--- program cerlaizgr (robot Fanuc LR Mate 200iD/7L) ---
  Suave(1)
  Establecer velocidad (1000.0 mm/s)
  Est. Ref.: bote cera
  Est. herr: Tool 1
  Mostrar Tool 1
  MoveJ 1 to (318.69, -45.69, 237.74) mm, rotated rx 168.3 ry -14.7 rz -86.98 deg; joints [83.928, 45.745, -7.693, -16.831, -73.362, 101.148]
  MoveL 2 to (318.69, -45.69, 237.74) mm, rotated rx 168.3 ry -14.7 rz -86.98 deg; joints [83.928, 45.745, -7.693, -16.831, -73.362, 101.148]
  MoveL 3 to (299.08, -45.69, 139.68) mm, rotated rx 168.3 ry -14.7 rz -86.98 deg; joints [84.076, 51.288, -16.777, -17.851, -64.646, 103.898]
  MoveL 4 to (299.08, -45.69, 139.68) mm, rotated rx 168.3 ry -14.7 rz -86.98 deg; joints [84.076, 51.288, -16.777, -17.851, -64.646, 103.898]
  Establecer velocidad (50.0 mm/s)
  MoveL 5 to (313.16, -44.5, 139.68) mm, rotated rx 168.3 ry -14.7 rz -86.98 deg; joints [83.886, 49.076, -18.597, -18.155, -62.971, 104.717]
  MoveL 6 to (327.32, -44.52, 139.68) mm, rotated rx 168.3 ry -14.7 rz -86.98 deg; joints [83.776, 46.952, -20.301, -18.453, -61.386, 105.433]
  MoveL 7 to (341.43, -45.73, 139.68) mm, rotated rx 168.3 ry -14.7 rz -86.98 deg; joints [83.752, 44.917, -21.892, -18.741, -59.886, 106.039]
  MoveL 8 to (355.34, -48.13, 139.68) mm, rotated rx 168.3 ry -14.7 rz -86.98 deg; joints [83.819, 42.973, -23.371, -19.018, -58.466, 106.529]
  MoveL 9 to (368.95, -51.69, 140.34) mm, rotated rx 168.3 ry -14.7 rz -86.98 deg; joints [83.98, 41.087, -24.673, -19.265, -57.187, 106.869]
  MoveL 10 to (383, -56.41, 142.33) mm, rotated rx 168.3 ry -14.7 rz -86.98 deg; joints [84.236, 39.118, -25.797, -19.475, -56.051, 107.053]
  MoveL 11 to (396.92, -60.57, 145.69) mm, rotated rx 168.3 ry -14.7 rz -86.98 deg; joints [84.459, 37.148, -26.671, -19.645, -55.16, 107.18]
  MoveL 12 to (410.7, -63.96, 150.39) mm, rotated rx 168.3 ry -14.7 rz -86.98 deg; joints [84.628, 35.164, -27.3, -19.771, -54.517, 107.266]
  MoveL 13 to (424.7, -66.68, 154.58) mm, rotated rx 168.3 ry -14.7 rz -86.98 deg; joints [84.746, 33.212, -27.925, -19.908, -53.893, 107.406]
  MoveL 14 to (439.04, -68.74, 157.38) mm, rotated rx 168.3 ry -14.7 rz -86.98 deg; joints [84.81, 31.317, -28.662, -20.086, -53.182, 107.653]
  MoveL 15 to (453.73, -70.09, 158.77) mm, rotated rx 168.3 ry -14.7 rz -86.98 deg; joints [84.812, 29.481, -29.518, -20.31, -52.377, 108.022]
  MoveL 16 to (469.71, -70.72, 158.92) mm, rotated rx 168.3 ry -14.7 rz -86.98 deg; joints [84.738, 27.589, -30.539, -20.6, -51.443, 108.552]
  MoveL 17 to (485.71, -70.47, 158.92) mm, rotated rx 168.3 ry -14.7 rz -86.98 deg; joints [84.58, 25.732, -31.509, -20.899, -50.584, 109.158]
  MoveL 18 to (501.7, -70.47, 158.92) mm, rotated rx 168.3 ry -14.7 rz -86.98 deg; joints [84.436, 23.886, -32.418, -21.19, -49.78, 109.731]
  MoveL 19 to (517.7, -70.47, 158.92) mm, rotated rx 168.3 ry -14.7 rz -86.98 deg; joints [84.284, 22.05, -33.266, -21.473, -49.036, 110.293]
  MoveL 20 to (533.69, -70.47, 158.92) mm, rotated rx 168.3 ry -14.7 rz -86.98 deg; joints [84.125, 20.219, -34.053, -21.748, -48.354, 110.844]
  MoveL 21 to (543.69, -70.47, 158.92) mm, rotated rx 168.3 ry -14.7 rz -86.98 deg; joints [84.02, 19.075, -34.514, -21.915, -47.958, 111.182]
  MoveL 22 to (553.68, -70.47, 158.92) mm, rotated rx 168.3 ry -14.7 rz -86.98 deg; joints [83.912, 17.931, -34.952, -22.077, -47.585, 111.515]
  MoveL 23 to (563.68, -70.47, 158.92) mm, rotated rx 168.3 ry -14.7 rz -86.98 deg; joints [83.799, 16.785, -35.366, -22.234, -47.237, 111.842]
  MoveL 24 to (573.77, -70.76, 158.92) mm, rotated rx 168.3 ry -14.7 rz -86.98 deg; joints [83.713, 15.622, -35.76, -22.383, -46.898, 112.135]
  MoveL 25 to (580.76, -72.49, 158.92) mm, rotated rx 168.3 ry -14.7 rz -86.98 deg; joints [83.817, 14.795, -36.025, -22.466, -46.622, 112.166]
  MoveL 26 to (587.5, -75.89, 158.92) mm, rotated rx 168.3 ry -14.7 rz -86.98 deg; joints [84.112, 13.973, -36.274, -22.521, -46.3, 111.995]
  MoveL 27 to (593.42, -80.86, 158.92) mm, rotated rx 168.3 ry -14.7 rz -86.98 deg; joints [84.6, 13.23, -36.489, -22.541, -45.951, 111.605]
  MoveL 28 to (598, -87.04, 158.92) mm, rotated rx 168.3 ry -14.7 rz -86.98 deg; joints [85.251, 12.632, -36.653, -22.52, -45.6, 111.02]
  MoveL 29 to (600.96, -93.88, 158.92) mm, rotated rx 168.3 ry -14.7 rz -86.98 deg; joints [86.003, 12.225, -36.76, -22.461, -45.269, 110.295]
  MoveL 30 to (602.27, -100.81, 158.92) mm, rotated rx 168.3 ry -14.7 rz -86.98 deg; joints [86.787, 12.02, -36.813, -22.373, -44.981, 109.505]
  MoveL 31 to (602.38, -107.49, 158.92) mm, rotated rx 168.3 ry -14.7 rz -86.98 deg; joints [87.553, 11.969, -36.826, -22.267, -44.736, 108.707]
  MoveL 32 to (602.38, -114.16, 158.92) mm, rotated rx 168.3 ry -14.7 rz -86.98 deg; joints [88.319, 11.941, -36.833, -22.154, -44.498, 107.903]
  MoveL 33 to (601.73, -120.97, 158.92) mm, rotated rx 168.3 ry -14.7 rz -86.98 deg; joints [89.103, 12, -36.818, -22.024, -44.276, 107.063]
  MoveL 34 to (599.51, -127.92, 158.92) mm, rotated rx 168.3 ry -14.7 rz -86.98 deg; joints [89.902, 12.254, -36.753, -21.866, -44.097, 106.177]
  MoveL 35 to (595.62, -134.46, 158.92) mm, rotated rx 168.3 ry -14.7 rz -86.98 deg; joints [90.646, 12.713, -36.63, -21.691, -43.99, 105.315]
  MoveL 36 to (590.24, -140.02, 158.92) mm, rotated rx 168.3 ry -14.7 rz -86.98 deg; joints [91.263, 13.353, -36.453, -21.513, -43.972, 104.557]
  MoveL 37 to (583.78, -144.14, 158.92) mm, rotated rx 168.3 ry -14.7 rz -86.98 deg; joints [91.703, 14.118, -36.231, -21.348, -44.05, 103.965]
  MoveL 38 to (576.83, -146.59, 158.92) mm, rotated rx 168.3 ry -14.7 rz -86.98 deg; joints [91.949, 14.935, -35.98, -21.209, -44.211, 103.569]
  MoveL 39 to (567.71, -147.44, 158.92) mm, rotated rx 168.3 ry -14.7 rz -86.98 deg; joints [92.006, 15.993, -35.636, -21.071, -44.515, 103.329]
  MoveL 40 to (558.83, -147.44, 158.92) mm, rotated rx 168.3 ry -14.7 rz -86.98 deg; joints [91.973, 17.018, -35.283, -20.949, -44.855, 103.185]
  MoveL 41 to (549.94, -147.44, 158.92) mm, rotated rx 168.3 ry -14.7 rz -86.98 deg; joints [91.941, 18.042, -34.91, -20.822, -45.212, 103.031]
  MoveL 42 to (541.06, -147.44, 158.92) mm, rotated rx 168.3 ry -14.7 rz -86.98 deg; joints [91.91, 19.064, -34.518, -20.691, -45.588, 102.87]
  MoveL 43 to (532.17, -147.44, 158.92) mm, rotated rx 168.3 ry -14.7 rz -86.98 deg; joints [91.88, 20.086, -34.107, -20.556, -45.981, 102.7]
  MoveL 44 to (523.28, -147.44, 158.92) mm, rotated rx 168.3 ry -14.7 rz -86.98 deg; joints [91.851, 21.107, -33.678, -20.417, -46.392, 102.523]
  MoveL 45 to (505.69, -147.44, 158.92) mm, rotated rx 168.3 ry -14.7 rz -86.98 deg; joints [91.796, 23.133, -32.772, -20.133, -47.257, 102.152]
  MoveL 46 to (488.1, -147.44, 158.92) mm, rotated rx 168.3 ry -14.7 rz -86.98 deg; joints [91.744, 25.167, -31.792, -19.839, -48.193, 101.755]
  MoveL 47 to (470.51, -148.03, 158.92) mm, rotated rx 168.3 ry -14.7 rz -86.98 deg; joints [91.749, 27.218, -30.736, -19.525, -49.186, 101.277]
  MoveL 48 to (453.01, -149.81, 158.74) mm, rotated rx 168.3 ry -14.7 rz -86.98 deg; joints [91.859, 29.295, -29.628, -19.193, -50.2, 100.677]
  MoveL 49 to (438.44, -152.23, 157.29) mm, rotated rx 168.3 ry -14.7 rz -86.98 deg; joints [92.027, 31.118, -28.792, -18.936, -50.942, 100.144]
  MoveL 50 to (424.24, -155.43, 154.47) mm, rotated rx 168.3 ry -14.7 rz -86.98 deg; joints [92.255, 32.993, -28.077, -18.707, -51.554, 99.605]
  MoveL 51 to (410.38, -159.2, 150.28) mm, rotated rx 168.3 ry -14.7 rz -86.98 deg; joints [92.522, 34.919, -27.475, -18.504, -52.049, 99.076]
  MoveL 52 to (396.59, -162.41, 145.59) mm, rotated rx 168.3 ry -14.7 rz -86.98 deg; joints [92.734, 36.883, -26.864, -18.314, -52.57, 98.606]
  MoveL 53 to (382.44, -164.94, 142.23) mm, rotated rx 168.3 ry -14.7 rz -86.98 deg; joints [92.881, 38.848, -26.002, -18.082, -53.348, 98.112]
  MoveL 54 to (367.94, -166.75, 140.25) mm, rotated rx 168.3 ry -14.7 rz -86.98 deg; joints [92.965, 40.825, -24.877, -17.812, -54.395, 97.593]
  MoveL 55 to (354.68, -167.73, 139.68) mm, rotated rx 168.3 ry -14.7 rz -86.98 deg; joints [92.987, 42.614, -23.639, -17.544, -55.567, 97.111]
  MoveL 56 to (341.32, -168.05, 139.68) mm, rotated rx 168.3 ry -14.7 rz -86.98 deg; joints [92.959, 44.442, -22.255, -17.273, -56.896, 96.643]
  MoveL 57 to (327.95, -168.05, 139.68) mm, rotated rx 168.3 ry -14.7 rz -86.98 deg; joints [92.908, 46.338, -20.784, -17.008, -58.316, 96.183]
  MoveL 58 to (314.6, -167.33, 139.68) mm, rotated rx 168.3 ry -14.7 rz -86.98 deg; joints [92.806, 48.311, -19.215, -16.755, -59.845, 95.759]
  MoveL 59 to (301.43, -165.08, 139.68) mm, rotated rx 168.3 ry -14.7 rz -86.98 deg; joints [92.599, 50.345, -17.557, -16.529, -61.49, 95.431]
  MoveL 60 to (288.61, -161.34, 139.93) mm, rotated rx 168.3 ry -14.7 rz -86.98 deg; joints [92.293, 52.424, -15.791, -16.327, -63.267, 95.183]
  MoveL 61 to (276.38, -156.17, 140.74) mm, rotated rx 168.3 ry -14.7 rz -86.98 deg; joints [91.9, 54.522, -13.891, -16.146, -65.197, 94.998]
  MoveL 62 to (264.77, -149.61, 142.03) mm, rotated rx 168.3 ry -14.7 rz -86.98 deg; joints [91.424, 56.664, -11.85, -15.987, -67.287, 94.869]
  MoveL 63 to (254.08, -141.83, 143.68) mm, rotated rx 168.3 ry -14.7 rz -86.98 deg; joints [90.88, 58.829, -9.702, -15.856, -69.499, 94.788]
  MoveL 64 to (248.15, -136.62, 144.8) mm, rotated rx 168.3 ry -14.7 rz -86.98 deg; joints [90.524, 60.146, -8.362, -15.79, -70.884, 94.76]
  MoveL 65 to (242.58, -131.01, 145.97) mm, rotated rx 168.3 ry -14.7 rz -86.98 deg; joints [90.146, 61.488, -6.978, -15.735, -72.318, 94.743]
  MoveL 66 to (237.41, -124.97, 147.17) mm, rotated rx 168.3 ry -14.7 rz -86.98 deg; joints [89.743, 62.855, -5.553, -15.69, -73.798, 94.742]
  MoveL 67 to (233.56, -118, 148.13) mm, rotated rx 168.3 ry -14.7 rz -86.98 deg; joints [89.284, 63.983, -4.368, -15.684, -75.063, 94.867]
  MoveL 68 to (231.55, -110.27, 148.66) mm, rotated rx 168.3 ry -14.7 rz -86.98 deg; joints [88.776, 64.645, -3.674, -15.726, -75.868, 95.177]
  MoveL 69 to (231.29, -101.33, 148.73) mm, rotated rx 168.3 ry -14.7 rz -86.98 deg; joints [88.187, 64.803, -3.515, -15.819, -76.181, 95.715]
  MoveL 70 to (231.99, -92.42, 148.54) mm, rotated rx 168.3 ry -14.7 rz -86.98 deg; joints [87.599, 64.684, -3.653, -15.931, -76.208, 96.336]
  MoveL 71 to (234.25, -83.83, 147.95) mm, rotated rx 168.3 ry -14.7 rz -86.98 deg; joints [87.025, 64.104, -4.279, -16.071, -75.764, 97.081]
  MoveL 72 to (237.98, -75.84, 147.03) mm, rotated rx 168.3 ry -14.7 rz -86.98 deg; joints [86.483, 63.146, -5.301, -16.236, -74.933, 97.911]
  MoveL 73 to (243.07, -68.63, 145.86) mm, rotated rx 168.3 ry -14.7 rz -86.98 deg; joints [85.983, 61.904, -6.611, -16.421, -73.816, 98.789]
  MoveL 74 to (249.32, -62.46, 144.57) mm, rotated rx 168.3 ry -14.7 rz -86.98 deg; joints [85.54, 60.474, -8.096, -16.619, -72.517, 99.67]
  MoveL 75 to (256.57, -57.48, 143.26) mm, rotated rx 168.3 ry -14.7 rz -86.98 deg; joints [85.167, 58.927, -9.672, -16.827, -71.114, 100.519]
  MoveL 76 to (264.6, -53.86, 142.05) mm, rotated rx 168.3 ry -14.7 rz -86.98 deg; joints [84.874, 57.321, -11.268, -17.037, -69.67, 101.305]
  MoveL 77 to (273.03, -51.14, 141.06) mm, rotated rx 168.3 ry -14.7 rz -86.98 deg; joints [84.635, 55.733, -12.799, -17.246, -68.277, 102.027]
  MoveL 78 to (281.59, -48.86, 140.32) mm, rotated rx 168.3 ry -14.7 rz -86.98 deg; joints [84.422, 54.21, -14.217, -17.452, -66.984, 102.699]
  MoveL 79 to (290.27, -47.04, 139.86) mm, rotated rx 168.3 ry -14.7 rz -86.98 deg; joints [84.235, 52.733, -15.54, -17.654, -65.778, 103.322]
  MoveL 80 to (299.08, -45.69, 139.68) mm, rotated rx 168.3 ry -14.7 rz -86.98 deg; joints [84.076, 51.288, -16.777, -17.851, -64.646, 103.898]
  Establecer velocidad (1000.0 mm/s)
  MoveL 81 to (299.08, -45.69, 139.68) mm, rotated rx 168.3 ry -14.7 rz -86.98 deg; joints [84.076, 51.288, -16.777, -17.851, -64.646, 103.898]
  MoveL 82 to (318.69, -45.69, 237.74) mm, rotated rx 168.3 ry -14.7 rz -86.98 deg; joints [83.928, 45.745, -7.693, -16.831, -73.362, 101.148]
  Establecer velocidad (1000.0 mm/s)
  MoveL 83 to (548.28, -147.66, 316.08) mm, rotated rx 168.3 ry -14.7 rz -86.98 deg; joints [91.957, 11.324, -13.989, -16.147, -65.087, 94.97]
  MoveL 84 to (528.67, -147.66, 218.02) mm, rotated rx 168.3 ry -14.7 rz -86.98 deg; joints [91.891, 17.173, -26.28, -18.338, -53.361, 99.273]
  MoveL 85 to (528.67, -147.66, 218.02) mm, rotated rx 168.3 ry -14.7 rz -86.98 deg; joints [91.891, 17.173, -26.28, -18.338, -53.361, 99.273]
  Establecer velocidad (50.0 mm/s)
  MoveL 86 to (522.32, -147.66, 218.02) mm, rotated rx 168.3 ry -14.7 rz -86.98 deg; joints [91.87, 17.943, -26.02, -18.282, -53.614, 99.193]
  MoveL 87 to (516.53, -147.66, 218.02) mm, rotated rx 168.3 ry -14.7 rz -86.98 deg; joints [91.851, 18.647, -25.772, -18.228, -53.854, 99.117]
  MoveL 88 to (511.92, -147.66, 218.02) mm, rotated rx 168.3 ry -14.7 rz -86.98 deg; joints [91.837, 19.208, -25.569, -18.185, -54.052, 99.054]
  MoveL 89 to (508.33, -147.66, 218.02) mm, rotated rx 168.3 ry -14.7 rz -86.98 deg; joints [91.825, 19.646, -25.406, -18.15, -54.209, 99.003]
  MoveL 90 to (504.19, -147.63, 218.02) mm, rotated rx 168.3 ry -14.7 rz -86.98 deg; joints [91.809, 20.15, -25.215, -18.111, -54.396, 98.947]
  MoveL 91 to (499.76, -147.37, 218.02) mm, rotated rx 168.3 ry -14.7 rz -86.98 deg; joints [91.772, 20.69, -25.005, -18.071, -54.605, 98.906]
  MoveL 92 to (494.1, -146.64, 218.02) mm, rotated rx 168.3 ry -14.7 rz -86.98 deg; joints [91.686, 21.379, -24.73, -18.027, -54.891, 98.892]
  MoveL 93 to (486.98, -145.04, 218.02) mm, rotated rx 168.3 ry -14.7 rz -86.98 deg; joints [91.517, 22.246, -24.373, -17.982, -55.279, 98.936]
  MoveL 94 to (480.5, -143.47, 218.02) mm, rotated rx 168.3 ry -14.7 rz -86.98 deg; joints [91.356, 23.038, -24.035, -17.941, -55.645, 98.979]
  MoveL 95 to (474.07, -142.24, 218.02) mm, rotated rx 168.3 ry -14.7 rz -86.98 deg; joints [91.229, 23.828, -23.689, -17.892, -56.01, 98.984]
  MoveL 96 to (467.53, -142.38, 218.02) mm, rotated rx 168.3 ry -14.7 rz -86.98 deg; joints [91.229, 24.638, -23.322, -17.816, -56.36, 98.849]
  MoveL 97 to (460.99, -142.59, 218.02) mm, rotated rx 168.3 ry -14.7 rz -86.98 deg; joints [91.235, 25.452, -22.943, -17.739, -56.719, 98.704]
  MoveL 98 to (454.45, -142.81, 218.02) mm, rotated rx 168.3 ry -14.7 rz -86.98 deg; joints [91.242, 26.27, -22.551, -17.66, -57.09, 98.554]
  MoveL 99 to (447.91, -142.98, 218.02) mm, rotated rx 168.3 ry -14.7 rz -86.98 deg; joints [91.245, 27.093, -22.147, -17.581, -57.475, 98.406]
  MoveL 100 to (442.07, -143.05, 218.02) mm, rotated rx 168.3 ry -14.7 rz -86.98 deg; joints [91.239, 27.832, -21.774, -17.511, -57.831, 98.279]
  MoveL 101 to (436.23, -142.98, 218.02) mm, rotated rx 168.3 ry -14.7 rz -86.98 deg; joints [91.223, 28.574, -21.392, -17.442, -58.201, 98.16]
  MoveL 102 to (430.39, -142.73, 218.02) mm, rotated rx 168.3 ry -14.7 rz -86.98 deg; joints [91.19, 29.32, -20.999, -17.376, -58.585, 98.057]
  MoveL 103 to (424.57, -142.19, 218.02) mm, rotated rx 168.3 ry -14.7 rz -86.98 deg; joints [91.135, 30.067, -20.597, -17.313, -58.984, 97.974]
  MoveL 104 to (418.82, -141.23, 218.02) mm, rotated rx 168.3 ry -14.7 rz -86.98 deg; joints [91.045, 30.811, -20.188, -17.258, -59.4, 97.927]
  MoveL 105 to (413.76, -138.38, 218.02) mm, rotated rx 168.3 ry -14.7 rz -86.98 deg; joints [90.799, 31.466, -19.822, -17.239, -59.818, 98.057]
  MoveL 106 to (409.91, -134.01, 218.02) mm, rotated rx 168.3 ry -14.7 rz -86.98 deg; joints [90.431, 31.965, -19.538, -17.258, -60.191, 98.341]
  MoveL 107 to (407.38, -128.76, 218.02) mm, rotated rx 168.3 ry -14.7 rz -86.98 deg; joints [89.996, 32.298, -19.348, -17.304, -60.495, 98.727]
  MoveL 108 to (406.69, -122.98, 218.02) mm, rotated rx 168.3 ry -14.7 rz -86.98 deg; joints [89.519, 32.391, -19.293, -17.379, -60.681, 99.202]
  MoveL 109 to (407.14, -120.09, 218.02) mm, rotated rx 168.3 ry -14.7 rz -86.98 deg; joints [89.279, 32.335, -19.326, -17.426, -60.718, 99.46]
  MoveL 110 to (407.92, -117.25, 218.02) mm, rotated rx 168.3 ry -14.7 rz -86.98 deg; joints [89.043, 32.238, -19.382, -17.477, -60.731, 99.723]
  MoveL 111 to (408.72, -114.41, 218.02) mm, rotated rx 168.3 ry -14.7 rz -86.98 deg; joints [88.807, 32.139, -19.439, -17.527, -60.744, 99.986]
  MoveL 112 to (409.54, -111.57, 218.02) mm, rotated rx 168.3 ry -14.7 rz -86.98 deg; joints [88.571, 32.04, -19.496, -17.577, -60.757, 100.25]
  MoveL 113 to (410.37, -108.75, 218.02) mm, rotated rx 168.3 ry -14.7 rz -86.98 deg; joints [88.334, 31.94, -19.553, -17.626, -60.77, 100.513]
  MoveL 114 to (411.04, -105.93, 218.02) mm, rotated rx 168.3 ry -14.7 rz -86.98 deg; joints [88.099, 31.864, -19.596, -17.673, -60.796, 100.77]
  MoveL 115 to (408.87, -99.66, 218.02) mm, rotated rx 168.3 ry -14.7 rz -86.98 deg; joints [87.586, 32.18, -19.415, -17.727, -61.115, 101.234]
  MoveL 116 to (406.88, -93.33, 218.02) mm, rotated rx 168.3 ry -14.7 rz -86.98 deg; joints [87.071, 32.482, -19.241, -17.781, -61.429, 101.701]
  MoveL 117 to (406.79, -88.92, 218.02) mm, rotated rx 168.3 ry -14.7 rz -86.98 deg; joints [86.708, 32.526, -19.216, -17.834, -61.558, 102.063]
  MoveL 118 to (408.24, -84.75, 218.02) mm, rotated rx 168.3 ry -14.7 rz -86.98 deg; joints [86.357, 32.368, -19.307, -17.905, -61.573, 102.454]
  MoveL 119 to (410.89, -81.21, 218.02) mm, rotated rx 168.3 ry -14.7 rz -86.98 deg; joints [86.05, 32.05, -19.49, -17.983, -61.487, 102.831]
  MoveL 120 to (415.2, -78.14, 218.02) mm, rotated rx 168.3 ry -14.7 rz -86.98 deg; joints [85.771, 31.513, -19.796, -18.077, -61.278, 103.224]
  MoveL 121 to (420.33, -76.88, 218.02) mm, rotated rx 168.3 ry -14.7 rz -86.98 deg; joints [85.633, 30.856, -20.164, -18.161, -60.969, 103.495]
  MoveL 122 to (425.6, -76.36, 218.02) mm, rotated rx 168.3 ry -14.7 rz -86.98 deg; joints [85.555, 30.18, -20.536, -18.237, -60.638, 103.708]
  MoveL 123 to (430.88, -76.05, 218.02) mm, rotated rx 168.3 ry -14.7 rz -86.98 deg; joints [85.494, 29.504, -20.901, -18.311, -60.309, 103.902]
  MoveL 124 to (436.16, -75.89, 218.02) mm, rotated rx 168.3 ry -14.7 rz -86.98 deg; joints [85.445, 28.83, -21.258, -18.383, -59.985, 104.082]
  MoveL 125 to (447.8, -75.87, 218.02) mm, rotated rx 168.3 ry -14.7 rz -86.98 deg; joints [85.362, 27.357, -22.015, -18.536, -59.291, 104.444]
  MoveL 126 to (459.44, -76.04, 218.02) mm, rotated rx 168.3 ry -14.7 rz -86.98 deg; joints [85.294, 25.897, -22.732, -18.683, -58.632, 104.781]
  MoveL 127 to (471.07, -76.17, 218.02) mm, rotated rx 168.3 ry -14.7 rz -86.98 deg; joints [85.219, 24.452, -23.408, -18.828, -58.014, 105.113]
  MoveL 128 to (482.52, -74.36, 218.02) mm, rotated rx 168.3 ry -14.7 rz -86.98 deg; joints [84.965, 23.061, -24.026, -18.992, -57.505, 105.61]
  MoveL 129 to (494.01, -72.39, 218.02) mm, rotated rx 168.3 ry -14.7 rz -86.98 deg; joints [84.685, 21.676, -24.61, -19.154, -57.036, 106.123]
  MoveL 130 to (505.68, -71.13, 218.02) mm, rotated rx 168.3 ry -14.7 rz -86.98 deg; joints [84.462, 20.271, -25.169, -19.305, -56.575, 106.572]
  MoveL 131 to (525.45, -70.42, 218.02) mm, rotated rx 168.3 ry -14.7 rz -86.98 deg; joints [84.203, 17.883, -26.041, -19.535, -55.83, 107.186]
  MoveL 132 to (545.24, -70.93, 218.02) mm, rotated rx 168.3 ry -14.7 rz -86.98 deg; joints [84.05, 15.486, -26.814, -19.734, -55.148, 107.657]
  MoveL 133 to (553.61, -71.56, 218.02) mm, rotated rx 168.3 ry -14.7 rz -86.98 deg; joints [84.024, 14.466, -27.111, -19.808, -54.876, 107.807]
  MoveL 134 to (561.96, -72.42, 218.02) mm, rotated rx 168.3 ry -14.7 rz -86.98 deg; joints [84.024, 13.445, -27.39, -19.875, -54.615, 107.923]
  MoveL 135 to (570.28, -73.54, 218.02) mm, rotated rx 168.3 ry -14.7 rz -86.98 deg; joints [84.051, 12.422, -27.649, -19.934, -54.363, 108.003]
  MoveL 136 to (578.56, -74.92, 218.02) mm, rotated rx 168.3 ry -14.7 rz -86.98 deg; joints [84.107, 11.399, -27.888, -19.986, -54.121, 108.047]
  MoveL 137 to (586.53, -77.56, 218.02) mm, rotated rx 168.3 ry -14.7 rz -86.98 deg; joints [84.307, 10.395, -28.104, -20.012, -53.858, 107.932]
  MoveL 138 to (593.61, -82.03, 218.02) mm, rotated rx 168.3 ry -14.7 rz -86.98 deg; joints [84.729, 9.477, -28.284, -20, -53.561, 107.575]
  MoveL 139 to (598.22, -86.42, 218.02) mm, rotated rx 168.3 ry -14.7 rz -86.98 deg; joints [85.179, 8.864, -28.395, -19.966, -53.322, 107.16]
  MoveL 140 to (601.98, -91.51, 218.02) mm, rotated rx 168.3 ry -14.7 rz -86.98 deg; joints [85.724, 8.35, -28.483, -19.911, -53.076, 106.634]
  MoveL 141 to (604.69, -97.29, 218.02) mm, rotated rx 168.3 ry -14.7 rz -86.98 deg; joints [86.365, 7.967, -28.545, -19.833, -52.826, 105.996]
  MoveL 142 to (606.15, -103.46, 218.02) mm, rotated rx 168.3 ry -14.7 rz -86.98 deg; joints [87.067, 7.742, -28.58, -19.736, -52.584, 105.282]
  MoveL 143 to (606.38, -109.87, 218.02) mm, rotated rx 168.3 ry -14.7 rz -86.98 deg; joints [87.809, 7.678, -28.589, -19.622, -52.356, 104.513]
  MoveL 144 to (605.62, -117.86, 218.02) mm, rotated rx 168.3 ry -14.7 rz -86.98 deg; joints [88.736, 7.743, -28.579, -19.468, -52.093, 103.538]
  MoveL 145 to (602.67, -125.36, 218.02) mm, rotated rx 168.3 ry -14.7 rz -86.98 deg; joints [89.607, 8.095, -28.524, -19.306, -51.891, 102.599]
  MoveL 146 to (597.87, -131.88, 218.02) mm, rotated rx 168.3 ry -14.7 rz -86.98 deg; joints [90.353, 8.688, -28.425, -19.15, -51.768, 101.769]
  MoveL 147 to (591.74, -137.15, 218.02) mm, rotated rx 168.3 ry -14.7 rz -86.98 deg; joints [90.943, 9.451, -28.288, -19.008, -51.728, 101.087]
  MoveL 148 to (584.66, -140.98, 218.02) mm, rotated rx 168.3 ry -14.7 rz -86.98 deg; joints [91.356, 10.331, -28.116, -18.888, -51.773, 100.579]
  MoveL 149 to (576.86, -143.14, 218.02) mm, rotated rx 168.3 ry -14.7 rz -86.98 deg; joints [91.572, 11.293, -27.911, -18.795, -51.905, 100.265]
  MoveL 150 to (552.86, -146.5, 218.02) mm, rotated rx 168.3 ry -14.7 rz -86.98 deg; joints [91.854, 14.231, -27.176, -18.56, -52.521, 99.668]
  MoveL 151 to (528.67, -147.66, 218.02) mm, rotated rx 168.3 ry -14.7 rz -86.98 deg; joints [91.891, 17.173, -26.28, -18.338, -53.361, 99.273]
  Establecer velocidad (1000.0 mm/s)
  MoveL 152 to (528.67, -147.66, 218.02) mm, rotated rx 168.3 ry -14.7 rz -86.98 deg; joints [91.891, 17.173, -26.28, -18.338, -53.361, 99.273]
  MoveL 153 to (548.28, -147.66, 316.08) mm, rotated rx 168.3 ry -14.7 rz -86.98 deg; joints [91.957, 11.324, -13.989, -16.147, -65.087, 94.97]

--- program cerladergr (robot Fanuc LR Mate 200iD/7L) ---
  Suave(1)
  Establecer velocidad (1000.0 mm/s)
  Est. Ref.: RobotiQ 2F-140 Gripper (Mechanism) Base
  Est. herr: Tool 1
  Mostrar Tool 1
  MoveJ 1 to (373, 259.19, 228.55) mm, rotated rx 167 ry -29.36 rz -83.53 deg; joints [63.32, 52.446, -7.256, -31.558, -87.99, 122.337]
  MoveL 2 to (373, 259.19, 228.55) mm, rotated rx 167 ry -29.36 rz -83.53 deg; joints [63.32, 52.446, -7.256, -31.558, -87.99, 122.337]
  MoveL 3 to (353.39, 259.19, 130.49) mm, rotated rx 167 ry -29.36 rz -83.53 deg; joints [63.923, 58.146, -15.764, -32.083, -80.447, 126.338]
  MoveL 4 to (353.39, 259.19, 130.49) mm, rotated rx 167 ry -29.36 rz -83.53 deg; joints [63.923, 58.146, -15.764, -32.083, -80.447, 126.338]
  Establecer velocidad (50.0 mm/s)
  MoveL 5 to (367.29, 260.82, 130.49) mm, rotated rx 167 ry -29.36 rz -83.53 deg; joints [63.398, 56.026, -17.663, -32.191, -79.106, 127.797]
  MoveL 6 to (381.28, 261, 130.49) mm, rotated rx 167 ry -29.36 rz -83.53 deg; joints [62.945, 53.943, -19.497, -32.321, -77.784, 129.167]
  MoveL 7 to (395.26, 260.88, 130.49) mm, rotated rx 167 ry -29.36 rz -83.53 deg; joints [62.498, 51.972, -21.202, -32.454, -76.569, 130.467]
  MoveL 8 to (409.21, 260.11, 130.72) mm, rotated rx 167 ry -29.36 rz -83.53 deg; joints [62.079, 50.06, -22.793, -32.592, -75.435, 131.686]
  MoveL 9 to (423.7, 258.54, 132.26) mm, rotated rx 167 ry -29.36 rz -83.53 deg; joints [61.68, 48.054, -24.243, -32.726, -74.413, 132.815]
  MoveL 10 to (437.83, 256.25, 135.18) mm, rotated rx 167 ry -29.36 rz -83.53 deg; joints [61.328, 46.053, -25.448, -32.843, -73.572, 133.774]
  MoveL 11 to (451.61, 253.27, 139.46) mm, rotated rx 167 ry -29.36 rz -83.53 deg; joints [61.022, 44.039, -26.42, -32.937, -72.906, 134.566]
  MoveL 12 to (465.25, 249.6, 144.01) mm, rotated rx 167 ry -29.36 rz -83.53 deg; joints [60.756, 42.031, -27.297, -33.029, -72.3, 135.274]
  MoveL 13 to (479.23, 246.21, 147.22) mm, rotated rx 167 ry -29.36 rz -83.53 deg; joints [60.449, 40.113, -28.251, -33.13, -71.648, 136.062]
  MoveL 14 to (493.56, 243.58, 149.07) mm, rotated rx 167 ry -29.36 rz -83.53 deg; joints [60.061, 38.316, -29.274, -33.229, -70.978, 136.953]
  MoveL 15 to (509.27, 241.65, 149.54) mm, rotated rx 167 ry -29.36 rz -83.53 deg; joints [59.551, 36.534, -30.453, -33.333, -70.236, 138.031]
  MoveL 16 to (525.09, 240.69, 149.54) mm, rotated rx 167 ry -29.36 rz -83.53 deg; joints [58.942, 34.866, -31.586, -33.406, -69.576, 139.158]
  MoveL 17 to (540.95, 240.59, 149.54) mm, rotated rx 167 ry -29.36 rz -83.53 deg; joints [58.245, 33.283, -32.628, -33.439, -69.032, 140.299]
  MoveL 18 to (556.8, 240.59, 149.54) mm, rotated rx 167 ry -29.36 rz -83.53 deg; joints [57.51, 31.74, -33.612, -33.447, -68.55, 141.431]
  MoveL 19 to (572.65, 240.59, 149.54) mm, rotated rx 167 ry -29.36 rz -83.53 deg; joints [56.745, 30.227, -34.544, -33.432, -68.121, 142.553]
  MoveL 20 to (612.29, 240.59, 149.54) mm, rotated rx 167 ry -29.36 rz -83.53 deg; joints [54.685, 26.561, -36.664, -33.285, -67.272, 145.325]
  MoveL 21 to (619.05, 240.05, 149.54) mm, rotated rx 167 ry -29.36 rz -83.53 deg; joints [54.353, 25.916, -37.015, -33.26, -67.124, 145.775]
  MoveL 22 to (625.97, 237.97, 149.54) mm, rotated rx 167 ry -29.36 rz -83.53 deg; joints [54.126, 25.159, -37.418, -33.281, -66.886, 146.18]
  MoveL 23 to (632.52, 234.23, 149.54) mm, rotated rx 167 ry -29.36 rz -83.53 deg; joints [54.047, 24.331, -37.849, -33.357, -66.56, 146.495]
  MoveL 24 to (638.13, 228.99, 149.54) mm, rotated rx 167 ry -29.36 rz -83.53 deg; joints [54.141, 23.491, -38.274, -33.491, -66.164, 146.682]
  MoveL 25 to (642.31, 222.67, 149.54) mm, rotated rx 167 ry -29.36 rz -83.53 deg; joints [54.41, 22.709, -38.659, -33.675, -65.727, 146.723]
  MoveL 26 to (644.86, 215.81, 149.54) mm, rotated rx 167 ry -29.36 rz -83.53 deg; joints [54.826, 22.043, -38.979, -33.894, -65.282, 146.622]
  MoveL 27 to (645.81, 209, 149.54) mm, rotated rx 167 ry -29.36 rz -83.53 deg; joints [55.341, 21.528, -39.22, -34.127, -64.858, 146.406]
  MoveL 28 to (645.83, 202.39, 149.54) mm, rotated rx 167 ry -29.36 rz -83.53 deg; joints [55.901, 21.115, -39.41, -34.363, -64.457, 146.128]
  MoveL 29 to (645.8, 195.79, 149.54) mm, rotated rx 167 ry -29.36 rz -83.53 deg; joints [56.471, 20.712, -39.593, -34.601, -64.057, 145.841]
  MoveL 30 to (644.81, 188.97, 149.54) mm, rotated rx 167 ry -29.36 rz -83.53 deg; joints [57.122, 20.392, -39.736, -34.854, -63.654, 145.473]
  MoveL 31 to (642.22, 182.12, 149.54) mm, rotated rx 167 ry -29.36 rz -83.53 deg; joints [57.871, 20.228, -39.809, -35.119, -63.264, 144.992]
  MoveL 32 to (637.99, 175.81, 149.54) mm, rotated rx 167 ry -29.36 rz -83.53 deg; joints [58.666, 20.259, -39.795, -35.37, -62.924, 144.424]
  MoveL 33 to (632.35, 170.61, 149.54) mm, rotated rx 167 ry -29.36 rz -83.53 deg; joints [59.434, 20.497, -39.689, -35.583, -62.667, 143.814]
  MoveL 34 to (625.78, 166.92, 149.54) mm, rotated rx 167 ry -29.36 rz -83.53 deg; joints [60.11, 20.918, -39.5, -35.737, -62.517, 143.213]
  MoveL 35 to (617.87, 164.72, 149.54) mm, rotated rx 167 ry -29.36 rz -83.53 deg; joints [60.708, 21.556, -39.207, -35.831, -62.484, 142.596]
  MoveL 36 to (610.22, 164.38, 149.54) mm, rotated rx 167 ry -29.36 rz -83.53 deg; joints [61.117, 22.275, -38.868, -35.852, -62.573, 142.082]
  MoveL 37 to (602.67, 164.38, 149.54) mm, rotated rx 167 ry -29.36 rz -83.53 deg; joints [61.482, 23.005, -38.514, -35.853, -62.692, 141.589]
  MoveL 38 to (595.12, 164.38, 149.54) mm, rotated rx 167 ry -29.36 rz -83.53 deg; joints [61.839, 23.737, -38.15, -35.848, -62.824, 141.095]
  MoveL 39 to (587.57, 164.38, 149.54) mm, rotated rx 167 ry -29.36 rz -83.53 deg; joints [62.187, 24.473, -37.775, -35.836, -62.967, 140.598]
  MoveL 40 to (580.02, 164.38, 149.54) mm, rotated rx 167 ry -29.36 rz -83.53 deg; joints [62.528, 25.212, -37.39, -35.818, -63.122, 140.099]
  MoveL 41 to (572.47, 164.38, 149.54) mm, rotated rx 167 ry -29.36 rz -83.53 deg; joints [62.861, 25.955, -36.993, -35.793, -63.288, 139.598]
  MoveL 42 to (555.03, 164.38, 149.54) mm, rotated rx 167 ry -29.36 rz -83.53 deg; joints [63.602, 27.686, -36.034, -35.714, -63.718, 138.432]
  MoveL 43 to (537.59, 164.38, 149.54) mm, rotated rx 167 ry -29.36 rz -83.53 deg; joints [64.307, 29.44, -35.015, -35.605, -64.212, 137.252]
  MoveL 44 to (520.16, 164.64, 149.54) mm, rotated rx 167 ry -29.36 rz -83.53 deg; joints [64.956, 31.235, -33.925, -35.463, -64.787, 136.068]
  MoveL 45 to (502.72, 164.25, 149.52) mm, rotated rx 167 ry -29.36 rz -83.53 deg; joints [65.625, 33.033, -32.792, -35.315, -65.388, 134.842]
  MoveL 46 to (488.07, 163.1, 148.53) mm, rotated rx 167 ry -29.36 rz -83.53 deg; joints [66.227, 34.592, -31.921, -35.22, -65.805, 133.834]
  MoveL 47 to (473.76, 161.25, 146.14) mm, rotated rx 167 ry -29.36 rz -83.53 deg; joints [66.85, 36.19, -31.203, -35.168, -66.086, 132.906]
  MoveL 48 to (459.79, 158.73, 142.36) mm, rotated rx 167 ry -29.36 rz -83.53 deg; joints [67.489, 37.827, -30.629, -35.152, -66.239, 132.054]
  MoveL 49 to (446.12, 155.56, 137.58) mm, rotated rx 167 ry -29.36 rz -83.53 deg; joints [68.148, 39.485, -30.151, -35.16, -66.303, 131.246]
  MoveL 50 to (432.36, 151.65, 133.88) mm, rotated rx 167 ry -29.36 rz -83.53 deg; joints [68.842, 41.087, -29.513, -35.13, -66.478, 130.308]
  MoveL 51 to (418.49, 146.99, 131.54) mm, rotated rx 167 ry -29.36 rz -83.53 deg; joints [69.572, 42.626, -28.685, -35.054, -66.789, 129.221]
  MoveL 52 to (403.25, 142.71, 130.51) mm, rotated rx 167 ry -29.36 rz -83.53 deg; joints [70.289, 44.319, -27.514, -34.889, -67.387, 127.929]
  MoveL 53 to (387.61, 139.91, 130.49) mm, rotated rx 167 ry -29.36 rz -83.53 deg; joints [70.886, 46.135, -26.064, -34.642, -68.274, 126.564]
  MoveL 54 to (371.71, 138.61, 130.49) mm, rotated rx 167 ry -29.36 rz -83.53 deg; joints [71.361, 48.132, -24.434, -34.35, -69.374, 125.194]
  MoveL 55 to (355.76, 138.87, 130.49) mm, rotated rx 167 ry -29.36 rz -83.53 deg; joints [71.713, 50.307, -22.617, -34.023, -70.695, 123.824]
  MoveL 56 to (339.98, 140.64, 130.57) mm, rotated rx 167 ry -29.36 rz -83.53 deg; joints [71.945, 52.659, -20.599, -33.672, -72.251, 122.449]
  MoveL 57 to (330.3, 142.51, 130.98) mm, rotated rx 167 ry -29.36 rz -83.53 deg; joints [72.031, 54.207, -19.195, -33.44, -73.376, 121.567]
  MoveL 58 to (320.78, 144.94, 131.74) mm, rotated rx 167 ry -29.36 rz -83.53 deg; joints [72.075, 55.829, -17.661, -33.202, -74.636, 120.654]
  MoveL 59 to (311.42, 147.93, 132.83) mm, rotated rx 167 ry -29.36 rz -83.53 deg; joints [72.077, 57.548, -15.977, -32.962, -76.046, 119.702]
  MoveL 60 to (302.56, 152.03, 134.18) mm, rotated rx 167 ry -29.36 rz -83.53 deg; joints [71.997, 59.362, -14.151, -32.725, -77.622, 118.752]
  MoveL 61 to (294.68, 157.81, 135.64) mm, rotated rx 167 ry -29.36 rz -83.53 deg; joints [71.791, 61.254, -12.215, -32.5, -79.36, 117.859]
  MoveL 62 to (288.13, 165, 137.04) mm, rotated rx 167 ry -29.36 rz -83.53 deg; joints [71.473, 63.168, -10.244, -32.302, -81.192, 117.055]
  MoveL 63 to (283.08, 173.42, 138.24) mm, rotated rx 167 ry -29.36 rz -83.53 deg; joints [71.053, 65.063, -8.295, -32.139, -83.061, 116.36]
  MoveL 64 to (279.82, 182.65, 139.07) mm, rotated rx 167 ry -29.36 rz -83.53 deg; joints [70.551, 66.824, -6.501, -32.018, -84.846, 115.826]
  MoveL 65 to (278.68, 189.17, 139.37) mm, rotated rx 167 ry -29.36 rz -83.53 deg; joints [70.175, 67.87, -5.452, -31.96, -85.934, 115.587]
  MoveL 66 to (278.41, 195.78, 139.44) mm, rotated rx 167 ry -29.36 rz -83.53 deg; joints [69.777, 68.748, -4.592, -31.917, -86.874, 115.468]
  MoveL 67 to (278.52, 202.41, 139.42) mm, rotated rx 167 ry -29.36 rz -83.53 deg; joints [69.371, 69.577, -3.786, -31.884, -87.772, 115.386]
  MoveL 68 to (279.75, 208.85, 139.09) mm, rotated rx 167 ry -29.36 rz -83.53 deg; joints [68.953, 70.031, -3.386, -31.863, -88.332, 115.529]
  MoveL 69 to (283.41, 216.79, 138.16) mm, rotated rx 167 ry -29.36 rz -83.53 deg; joints [68.387, 69.813, -3.726, -31.847, -88.341, 116.188]
  MoveL 70 to (288.89, 223.57, 136.87) mm, rotated rx 167 ry -29.36 rz -83.53 deg; joints [67.847, 68.844, -4.849, -31.843, -87.671, 117.239]
  MoveL 71 to (294.97, 229.75, 135.58) mm, rotated rx 167 ry -29.36 rz -83.53 deg; joints [67.324, 67.735, -6.1, -31.845, -86.883, 118.343]
  MoveL 72 to (304.9, 238.1, 133.79) mm, rotated rx 167 ry -29.36 rz -83.53 deg; joints [66.567, 65.979, -8.03, -31.86, -85.641, 120.003]
  MoveL 73 to (315.82, 245.35, 132.28) mm, rotated rx 167 ry -29.36 rz -83.53 deg; joints [65.839, 64.126, -9.995, -31.891, -84.351, 121.657]
  MoveL 74 to (327.51, 251.3, 131.17) mm, rotated rx 167 ry -29.36 rz -83.53 deg; joints [65.156, 62.215, -11.938, -31.937, -83.057, 123.263]
  MoveL 75 to (339.8, 255.89, 130.57) mm, rotated rx 167 ry -29.36 rz -83.53 deg; joints [64.527, 60.262, -13.825, -31.999, -81.78, 124.796]
  Establecer velocidad (1000.0 mm/s)
  MoveL 76 to (339.8, 255.89, 130.57) mm, rotated rx 167 ry -29.36 rz -83.53 deg; joints [64.527, 60.262, -13.825, -31.999, -81.78, 124.796]
  MoveL 77 to (359.41, 255.89, 228.63) mm, rotated rx 167 ry -29.36 rz -83.53 deg; joints [63.945, 54.713, -5.34, -31.591, -89.297, 120.804]
  Establecer velocidad (1000.0 mm/s)
  MoveL 78 to (592.45, 240.79, 306.28) mm, rotated rx 167 ry -29.36 rz -83.53 deg; joints [55.727, 21.015, -16.141, -30.759, -84.238, 133.32]
  MoveL 79 to (572.84, 240.79, 208.22) mm, rotated rx 167 ry -29.36 rz -83.53 deg; joints [56.72, 26.836, -27.528, -32.122, -74.034, 138.559]
  MoveL 80 to (572.84, 240.79, 208.22) mm, rotated rx 167 ry -29.36 rz -83.53 deg; joints [56.72, 26.836, -27.528, -32.122, -74.034, 138.559]
  Establecer velocidad (50.0 mm/s)
  MoveL 81 to (596.66, 239.65, 208.22) mm, rotated rx 167 ry -29.36 rz -83.53 deg; joints [55.594, 24.393, -28.729, -32.021, -73.544, 140.099]
  MoveL 82 to (620.29, 236.36, 208.22) mm, rotated rx 167 ry -29.36 rz -83.53 deg; joints [54.572, 21.873, -29.865, -31.928, -73.052, 141.517]
  MoveL 83 to (627.98, 234.28, 208.22) mm, rotated rx 167 ry -29.36 rz -83.53 deg; joints [54.302, 20.992, -30.237, -31.914, -72.86, 141.929]
  MoveL 84 to (634.98, 230.57, 208.22) mm, rotated rx 167 ry -29.36 rz -83.53 deg; joints [54.197, 20.067, -30.612, -31.947, -72.59, 142.218]
  MoveL 85 to (641.07, 225.44, 208.22) mm, rotated rx 167 ry -29.36 rz -83.53 deg; joints [54.257, 19.133, -30.976, -32.025, -72.253, 142.375]
  MoveL 86 to (645.86, 219.11, 208.22) mm, rotated rx 167 ry -29.36 rz -83.53 deg; joints [54.494, 18.24, -31.31, -32.149, -71.863, 142.38]
  MoveL 87 to (648.89, 211.77, 208.22) mm, rotated rx 167 ry -29.36 rz -83.53 deg; joints [54.927, 17.45, -31.592, -32.321, -71.427, 142.21]
  MoveL 88 to (649.78, 203.89, 208.22) mm, rotated rx 167 ry -29.36 rz -83.53 deg; joints [55.543, 16.834, -31.805, -32.533, -70.966, 141.862]
  MoveL 89 to (649.4, 195.99, 208.22) mm, rotated rx 167 ry -29.36 rz -83.53 deg; joints [56.246, 16.35, -31.967, -32.759, -70.508, 141.423]
  MoveL 90 to (647.13, 188.46, 208.22) mm, rotated rx 167 ry -29.36 rz -83.53 deg; joints [57.034, 16.084, -32.054, -32.993, -70.072, 140.877]
  MoveL 91 to (642.97, 181.75, 208.22) mm, rotated rx 167 ry -29.36 rz -83.53 deg; joints [57.862, 16.073, -32.058, -33.218, -69.686, 140.253]
  MoveL 92 to (637.44, 176.12, 208.22) mm, rotated rx 167 ry -29.36 rz -83.53 deg; joints [58.668, 16.279, -31.99, -33.418, -69.367, 139.604]
  MoveL 93 to (631.03, 171.89, 208.22) mm, rotated rx 167 ry -29.36 rz -83.53 deg; joints [59.389, 16.669, -31.86, -33.579, -69.137, 138.981]
  MoveL 94 to (623.86, 169.18, 208.22) mm, rotated rx 167 ry -29.36 rz -83.53 deg; joints [60.006, 17.238, -31.666, -33.696, -69.009, 138.399]
  MoveL 95 to (616.37, 167.81, 208.22) mm, rotated rx 167 ry -29.36 rz -83.53 deg; joints [60.508, 17.924, -31.424, -33.77, -68.973, 137.874]
  MoveL 96 to (608.82, 166.72, 208.22) mm, rotated rx 167 ry -29.36 rz -83.53 deg; joints [60.979, 18.636, -31.163, -33.83, -68.965, 137.36]
  MoveL 97 to (589.49, 164.88, 208.22) mm, rotated rx 167 ry -29.36 rz -83.53 deg; joints [62.056, 20.534, -30.424, -33.929, -69.063, 136.096]
  MoveL 98 to (570.08, 164.36, 208.22) mm, rotated rx 167 ry -29.36 rz -83.53 deg; joints [62.967, 22.539, -29.574, -33.955, -69.327, 134.889]
  MoveL 99 to (552.43, 164.88, 208.22) mm, rotated rx 167 ry -29.36 rz -83.53 deg; joints [63.668, 24.438, -28.707, -33.926, -69.705, 133.829]
  MoveL 100 to (534.96, 166.82, 208.22) mm, rotated rx 167 ry -29.36 rz -83.53 deg; joints [64.211, 26.415, -27.741, -33.842, -70.24, 132.833]
  MoveL 101 to (517.84, 170.06, 208.22) mm, rotated rx 167 ry -29.36 rz -83.53 deg; joints [64.61, 28.451, -26.682, -33.713, -70.923, 131.896]
  MoveL 102 to (500.39, 169.87, 208.22) mm, rotated rx 167 ry -29.36 rz -83.53 deg; joints [65.267, 30.376, -25.621, -33.635, -71.479, 130.756]
  MoveL 103 to (482.95, 169.78, 208.22) mm, rotated rx 167 ry -29.36 rz -83.53 deg; joints [65.887, 32.348, -24.479, -33.536, -72.12, 129.599]
  MoveL 104 to (477.76, 169.9, 208.22) mm, rotated rx 167 ry -29.36 rz -83.53 deg; joints [66.054, 32.952, -24.119, -33.5, -72.336, 129.256]
  MoveL 105 to (472.58, 170.16, 208.22) mm, rotated rx 167 ry -29.36 rz -83.53 deg; joints [66.209, 33.566, -23.747, -33.461, -72.568, 128.917]
  MoveL 106 to (467.41, 170.6, 208.22) mm, rotated rx 167 ry -29.36 rz -83.53 deg; joints [66.347, 34.193, -23.361, -33.417, -72.82, 128.584]
  MoveL 107 to (462.3, 171.44, 208.22) mm, rotated rx 167 ry -29.36 rz -83.53 deg; joints [66.452, 34.838, -22.959, -33.366, -73.103, 128.268]
  MoveL 108 to (457.78, 173.91, 208.22) mm, rotated rx 167 ry -29.36 rz -83.53 deg; joints [66.415, 35.504, -22.538, -33.291, -73.474, 128.057]
  MoveL 109 to (454.83, 177.06, 208.22) mm, rotated rx 167 ry -29.36 rz -83.53 deg; joints [66.277, 36.022, -22.206, -33.216, -73.821, 127.979]
  MoveL 110 to (452.9, 180.92, 208.22) mm, rotated rx 167 ry -29.36 rz -83.53 deg; joints [66.056, 36.458, -21.924, -33.138, -74.169, 127.996]
  MoveL 111 to (452.35, 185.18, 208.22) mm, rotated rx 167 ry -29.36 rz -83.53 deg; joints [65.762, 36.755, -21.731, -33.063, -74.48, 128.124]
  MoveL 112 to (453.25, 189.41, 208.22) mm, rotated rx 167 ry -29.36 rz -83.53 deg; joints [65.425, 36.878, -21.651, -32.999, -74.718, 128.351]
  MoveL 113 to (454.63, 193.53, 208.22) mm, rotated rx 167 ry -29.36 rz -83.53 deg; joints [65.079, 36.94, -21.61, -32.938, -74.927, 128.607]
  MoveL 114 to (456.04, 197.65, 208.22) mm, rotated rx 167 ry -29.36 rz -83.53 deg; joints [64.734, 37.002, -21.57, -32.878, -75.135, 128.863]
  MoveL 115 to (456.44, 200.94, 208.22) mm, rotated rx 167 ry -29.36 rz -83.53 deg; joints [64.484, 37.142, -21.477, -32.824, -75.339, 129.014]
  MoveL 116 to (455.45, 204.28, 208.22) mm, rotated rx 167 ry -29.36 rz -83.53 deg; joints [64.279, 37.454, -21.272, -32.762, -75.616, 129.065]
  MoveL 117 to (454.48, 207.62, 208.22) mm, rotated rx 167 ry -29.36 rz -83.53 deg; joints [64.073, 37.765, -21.065, -32.7, -75.893, 129.115]
  MoveL 118 to (453.53, 210.97, 208.22) mm, rotated rx 167 ry -29.36 rz -83.53 deg; joints [63.869, 38.078, -20.856, -32.639, -76.172, 129.165]
  MoveL 119 to (452.65, 214.33, 208.22) mm, rotated rx 167 ry -29.36 rz -83.53 deg; joints [63.662, 38.385, -20.649, -32.579, -76.45, 129.219]
  MoveL 120 to (452.59, 220.11, 208.22) mm, rotated rx 167 ry -29.36 rz -83.53 deg; joints [63.258, 38.744, -20.407, -32.482, -76.858, 129.412]
  MoveL 121 to (454.53, 225.57, 208.22) mm, rotated rx 167 ry -29.36 rz -83.53 deg; joints [62.808, 38.846, -20.338, -32.399, -77.143, 129.74]
  MoveL 122 to (457.95, 230.26, 208.22) mm, rotated rx 167 ry -29.36 rz -83.53 deg; joints [62.358, 38.726, -20.419, -32.333, -77.299, 130.149]
  MoveL 123 to (461.85, 233.35, 208.22) mm, rotated rx 167 ry -29.36 rz -83.53 deg; joints [62.001, 38.453, -20.604, -32.293, -77.322, 130.54]
  MoveL 124 to (466.6, 234.84, 208.22) mm, rotated rx 167 ry -29.36 rz -83.53 deg; joints [61.721, 37.981, -20.921, -32.282, -77.194, 130.941]
  MoveL 125 to (471.6, 235.51, 208.22) mm, rotated rx 167 ry -29.36 rz -83.53 deg; joints [61.486, 37.434, -21.285, -32.285, -77.003, 131.33]
  MoveL 126 to (476.62, 235.91, 208.22) mm, rotated rx 167 ry -29.36 rz -83.53 deg; joints [61.267, 36.873, -21.655, -32.291, -76.8, 131.71]
  MoveL 127 to (481.65, 236.12, 208.22) mm, rotated rx 167 ry -29.36 rz -83.53 deg; joints [61.058, 36.304, -22.025, -32.298, -76.591, 132.082]
  MoveL 128 to (486.68, 236.18, 208.22) mm, rotated rx 167 ry -29.36 rz -83.53 deg; joints [60.857, 35.732, -22.393, -32.308, -76.379, 132.446]
  MoveL 129 to (491.7, 236.14, 208.22) mm, rotated rx 167 ry -29.36 rz -83.53 deg; joints [60.661, 35.159, -22.757, -32.317, -76.168, 132.804]
  MoveL 130 to (502.02, 235.87, 208.22) mm, rotated rx 167 ry -29.36 rz -83.53 deg; joints [60.263, 33.986, -23.489, -32.336, -75.745, 133.526]
  MoveL 131 to (512.35, 235.54, 208.22) mm, rotated rx 167 ry -29.36 rz -83.53 deg; joints [59.86, 32.829, -24.193, -32.351, -75.347, 134.237]
  MoveL 132 to (522.6, 236.12, 208.22) mm, rotated rx 167 ry -29.36 rz -83.53 deg; joints [59.382, 31.755, -24.83, -32.34, -75.042, 134.969]
  MoveL 133 to (532.92, 238.55, 208.22) mm, rotated rx 167 ry -29.36 rz -83.53 deg; joints [58.754, 30.809, -25.376, -32.281, -74.884, 135.769]
  MoveL 134 to (539.18, 239.87, 208.22) mm, rotated rx 167 ry -29.36 rz -83.53 deg; joints [58.377, 30.234, -25.702, -32.243, -74.79, 136.247]
  MoveL 135 to (544.13, 240.49, 208.22) mm, rotated rx 167 ry -29.36 rz -83.53 deg; joints [58.106, 29.757, -25.969, -32.22, -74.694, 136.609]
  MoveL 136 to (547.94, 240.73, 208.22) mm, rotated rx 167 ry -29.36 rz -83.53 deg; joints [57.913, 29.376, -26.18, -32.207, -74.609, 136.878]
  MoveL 137 to (551.23, 240.79, 208.22) mm, rotated rx 167 ry -29.36 rz -83.53 deg; joints [57.756, 29.039, -26.364, -32.197, -74.528, 137.103]
  MoveL 138 to (554.67, 240.79, 208.22) mm, rotated rx 167 ry -29.36 rz -83.53 deg; joints [57.595, 28.685, -26.556, -32.188, -74.442, 137.335]
  MoveL 139 to (558, 240.79, 208.22) mm, rotated rx 167 ry -29.36 rz -83.53 deg; joints [57.438, 28.343, -26.74, -32.178, -74.361, 137.56]
  MoveL 140 to (562.29, 240.79, 208.22) mm, rotated rx 167 ry -29.36 rz -83.53 deg; joints [57.233, 27.905, -26.973, -32.163, -74.261, 137.85]
  MoveL 141 to (567.43, 240.79, 208.22) mm, rotated rx 167 ry -29.36 rz -83.53 deg; joints [56.985, 27.382, -27.246, -32.144, -74.148, 138.196]
  MoveL 142 to (572.84, 240.79, 208.22) mm, rotated rx 167 ry -29.36 rz -83.53 deg; joints [56.72, 26.836, -27.528, -32.122, -74.034, 138.559]
  Establecer velocidad (1000.0 mm/s)
  MoveL 143 to (572.84, 240.79, 208.22) mm, rotated rx 167 ry -29.36 rz -83.53 deg; joints [56.72, 26.836, -27.528, -32.122, -74.034, 138.559]
  MoveL 144 to (592.45, 240.79, 306.28) mm, rotated rx 167 ry -29.36 rz -83.53 deg; joints [55.727, 21.015, -16.141, -30.759, -84.238, 133.32]

--- program ceraariizgr (robot Fanuc LR Mate 200iD/7L) ---
  Suave(1)
  Establecer velocidad (1000.0 mm/s)
  Est. Ref.: RobotiQ 2F-140 Gripper (Mechanism) Base
  Est. herr: Tool 1
  Mostrar Tool 1
  MoveJ 1 to (325.94, -36.21, 264.31) mm, rotated rx 167.98 ry -19.59 rz -85.91 deg; joints [81.562, 45.316, -5.344, -21.983, -77.448, 103.906]
  MoveL 2 to (325.94, -36.21, 264.31) mm, rotated rx 167.98 ry -19.59 rz -85.91 deg; joints [81.562, 45.316, -5.344, -21.983, -77.448, 103.906]
  MoveL 3 to (306.33, -36.21, 166.25) mm, rotated rx 167.98 ry -19.59 rz -85.91 deg; joints [81.767, 50.338, -14.842, -23.076, -68.594, 107.512]
  MoveL 4 to (306.33, -36.21, 166.25) mm, rotated rx 167.98 ry -19.59 rz -85.91 deg; joints [81.767, 50.338, -14.842, -23.076, -68.594, 107.512]
  Establecer velocidad (50.0 mm/s)
  MoveL 5 to (294.66, -36.21, 164.87) mm, rotated rx 167.98 ry -19.59 rz -85.91 deg; joints [81.884, 52.376, -13.349, -22.844, -69.925, 106.778]
  MoveL 6 to (282.99, -36.21, 163.24) mm, rotated rx 167.98 ry -19.59 rz -85.91 deg; joints [81.999, 54.551, -11.731, -22.613, -71.374, 106.006]
  MoveL 7 to (270.07, -36.21, 161.14) mm, rotated rx 167.98 ry -19.59 rz -85.91 deg; joints [82.121, 57.167, -9.745, -22.358, -73.162, 105.092]
  MoveL 8 to (255.49, -36.21, 158.4) mm, rotated rx 167.98 ry -19.59 rz -85.91 deg; joints [82.255, 60.494, -7.141, -22.067, -75.523, 103.942]
  MoveL 9 to (242.99, -36.21, 155.72) mm, rotated rx 167.98 ry -19.59 rz -85.91 deg; joints [82.366, 63.851, -4.405, -21.814, -78.02, 102.787]
  MoveL 10 to (237.07, -36.21, 154.35) mm, rotated rx 167.98 ry -19.59 rz -85.91 deg; joints [82.418, 65.714, -2.831, -21.691, -79.463, 102.143]
  MoveL 11 to (231.82, -36.21, 153.08) mm, rotated rx 167.98 ry -19.59 rz -85.91 deg; joints [82.463, 67.62, -1.176, -21.581, -80.985, 101.482]
  MoveL 12 to (229.61, -36.21, 152.44) mm, rotated rx 167.98 ry -19.59 rz -85.91 deg; joints [82.482, 68.523, -0.386, -21.534, -81.712, 101.17]
  MoveL 13 to (228.19, -36.21, 151.51) mm, rotated rx 167.98 ry -19.59 rz -85.91 deg; joints [82.494, 69.131, 0.081, -21.508, -82.143, 100.986]
  MoveL 14 to (226.98, -36.21, 149.94) mm, rotated rx 167.98 ry -19.59 rz -85.91 deg; joints [82.504, 69.641, 0.367, -21.493, -82.405, 100.871]
  MoveL 15 to (226.47, -36.21, 148.43) mm, rotated rx 167.98 ry -19.59 rz -85.91 deg; joints [82.509, 69.827, 0.344, -21.493, -82.382, 100.875]
  MoveL 16 to (226.38, -36.21, 146.6) mm, rotated rx 167.98 ry -19.59 rz -85.91 deg; joints [82.509, 69.793, 0.061, -21.507, -82.118, 100.979]
  MoveL 17 to (226.38, -36.21, 144.11) mm, rotated rx 167.98 ry -19.59 rz -85.91 deg; joints [82.509, 69.697, -0.373, -21.53, -81.715, 101.14]
  MoveL 18 to (226.38, -36.21, 139.71) mm, rotated rx 167.98 ry -19.59 rz -85.91 deg; joints [82.509, 69.554, -1.114, -21.571, -81.026, 101.415]
  MoveL 19 to (226.38, -36.21, 134.59) mm, rotated rx 167.98 ry -19.59 rz -85.91 deg; joints [82.509, 69.427, -1.934, -21.621, -80.263, 101.721]
  MoveL 20 to (226.38, -36.21, 129.47) mm, rotated rx 167.98 ry -19.59 rz -85.91 deg; joints [82.509, 69.336, -2.72, -21.673, -79.532, 102.015]
  MoveL 21 to (226.38, -36.21, 124.22) mm, rotated rx 167.98 ry -19.59 rz -85.91 deg; joints [82.509, 69.276, -3.494, -21.727, -78.813, 102.307]
  Establecer velocidad (1000.0 mm/s)
  MoveL 22 to (226.38, -36.21, 124.22) mm, rotated rx 167.98 ry -19.59 rz -85.91 deg; joints [82.509, 69.276, -3.494, -21.727, -78.813, 102.307]
  MoveL 23 to (245.99, -36.21, 222.28) mm, rotated rx 167.98 ry -19.59 rz -85.91 deg; joints [82.34, 65.173, 5.951, -21.338, -87.663, 98.978]
  Establecer velocidad (1000.0 mm/s)
  MoveL 24 to (337.7, -36.21, 265.46) mm, rotated rx 167.98 ry -19.59 rz -85.91 deg; joints [81.434, 43.24, -6.701, -22.117, -76.237, 104.551]
  MoveL 25 to (318.09, -36.21, 167.4) mm, rotated rx 167.98 ry -19.59 rz -85.91 deg; joints [81.646, 48.398, -16.248, -23.311, -67.348, 108.226]
  MoveL 26 to (318.09, -36.21, 167.4) mm, rotated rx 167.98 ry -19.59 rz -85.91 deg; joints [81.646, 48.398, -16.248, -23.311, -67.348, 108.226]
  Establecer velocidad (50.0 mm/s)
  MoveL 27 to (340.29, -36.21, 170.42) mm, rotated rx 167.98 ry -19.59 rz -85.91 deg; joints [81.406, 44.926, -18.529, -23.73, -65.348, 109.449]
  MoveL 28 to (364.68, -36.21, 176.36) mm, rotated rx 167.98 ry -19.59 rz -85.91 deg; joints [81.126, 41.251, -20.404, -24.113, -63.741, 110.558]
  MoveL 29 to (388.28, -36.21, 184.92) mm, rotated rx 167.98 ry -19.59 rz -85.91 deg; joints [80.838, 37.74, -21.618, -24.385, -62.744, 111.391]
  MoveL 30 to (410.8, -36.21, 196.02) mm, rotated rx 167.98 ry -19.59 rz -85.91 deg; joints [80.545, 34.366, -22.209, -24.532, -62.319, 111.946]
  MoveL 31 to (431.97, -36.21, 209.51) mm, rotated rx 167.98 ry -19.59 rz -85.91 deg; joints [80.252, 31.132, -22.202, -24.549, -62.438, 112.221]
  MoveL 32 to (451.54, -36.21, 225.23) mm, rotated rx 167.98 ry -19.59 rz -85.91 deg; joints [79.964, 28.056, -21.624, -24.443, -63.074, 112.224]
  MoveL 33 to (469.27, -36.21, 242.99) mm, rotated rx 167.98 ry -19.59 rz -85.91 deg; joints [79.689, 25.178, -20.51, -24.232, -64.195, 111.973]
  Establecer velocidad (1000.0 mm/s)
  MoveL 34 to (469.27, -36.21, 242.99) mm, rotated rx 167.98 ry -19.59 rz -85.91 deg; joints [79.689, 25.178, -20.51, -24.232, -64.195, 111.973]
  MoveL 35 to (488.89, -36.21, 341.05) mm, rotated rx 167.98 ry -19.59 rz -85.91 deg; joints [79.366, 20.377, -8.926, -22.539, -74.958, 107.38]
  Establecer velocidad (1000.0 mm/s)
  MoveL 36 to (611.58, -36.21, 341.05) mm, rotated rx 167.98 ry -19.59 rz -85.91 deg; joints [76.791, 4.672, -12.49, -23.14, -72.655, 111.248]
  MoveL 37 to (591.97, -36.21, 242.99) mm, rotated rx 167.98 ry -19.59 rz -85.91 deg; joints [77.283, 10.263, -25.488, -25.437, -60.607, 116.6]
  MoveL 38 to (591.97, -36.21, 242.99) mm, rotated rx 167.98 ry -19.59 rz -85.91 deg; joints [77.283, 10.263, -25.488, -25.437, -60.607, 116.6]
  Establecer velocidad (50.0 mm/s)
  MoveL 39 to (599.82, -36.21, 201.76) mm, rotated rx 167.98 ry -19.59 rz -85.91 deg; joints [77.091, 11.534, -31.335, -27.056, -55.435, 119.826]
  MoveL 40 to (599.82, -36.21, 201.76) mm, rotated rx 167.98 ry -19.59 rz -85.91 deg; joints [77.091, 11.534, -31.335, -27.056, -55.435, 119.826]
  MoveL 41 to (602.6, -36.21, 182.64) mm, rotated rx 167.98 ry -19.59 rz -85.91 deg; joints [77.022, 12.423, -34.06, -27.962, -53.046, 121.441]
  MoveL 42 to (602.64, -36.21, 163.32) mm, rotated rx 167.98 ry -19.59 rz -85.91 deg; joints [77.021, 13.763, -36.744, -28.967, -50.686, 123.068]
  MoveL 43 to (599.94, -36.21, 144.19) mm, rotated rx 167.98 ry -19.59 rz -85.91 deg; joints [77.088, 15.506, -39.304, -30.044, -48.431, 124.664]
  MoveL 44 to (597.47, -36.21, 134.41) mm, rotated rx 167.98 ry -19.59 rz -85.91 deg; joints [77.15, 16.555, -40.561, -30.621, -47.323, 125.465]
  Establecer velocidad (1000.0 mm/s)
  MoveL 45 to (597.47, -36.21, 134.41) mm, rotated rx 167.98 ry -19.59 rz -85.91 deg; joints [77.15, 16.555, -40.561, -30.621, -47.323, 125.465]
  MoveL 46 to (617.08, -36.21, 232.47) mm, rotated rx 167.98 ry -19.59 rz -85.91 deg; joints [76.648, 7.748, -27.469, -25.951, -59.068, 118.186]

--- program cerarridergr (robot Fanuc LR Mate 200iD/7L) ---
  Suave(1)
  Establecer velocidad (1000.0 mm/s)
  Est. Ref.: RobotiQ 2F-140 Gripper (Mechanism) Base
  Est. herr: Tool 1
  Mostrar Tool 1
  MoveJ 1 to (442.77, 170.06, 192.98) mm, rotated rx 122.56 ry -24.48 rz -84.76 deg; joints [65.259, 23.707, -47.429, -101.449, -38.805, -167.89]
  MoveL 2 to (442.77, 170.06, 192.98) mm, rotated rx 122.56 ry -24.48 rz -84.76 deg; joints [65.259, 23.707, -47.429, -101.449, -38.805, -167.89]
  MoveL 3 to (423.16, 170.06, 94.92) mm, rotated rx 122.56 ry -24.48 rz -84.76 deg; joints [66.107, 35.403, -58.417, -114.705, -41.754, -151.456]
  MoveL 4 to (423.16, 170.06, 94.92) mm, rotated rx 122.56 ry -24.48 rz -84.76 deg; joints [66.107, 35.403, -58.417, -114.705, -41.754, -151.456]
  Establecer velocidad (50.0 mm/s)
  MoveL 5 to (420.64, 170.06, 94.69) mm, rotated rx 122.56 ry -24.48 rz -84.76 deg; joints [66.212, 35.616, -58.253, -114.653, -41.636, -151.645]
  MoveL 6 to (418.13, 170.06, 94.46) mm, rotated rx 122.56 ry -24.48 rz -84.76 deg; joints [66.316, 35.828, -58.088, -114.598, -41.517, -151.838]
  MoveL 7 to (411.73, 170.06, 93.82) mm, rotated rx 122.56 ry -24.48 rz -84.76 deg; joints [66.577, 36.378, -57.67, -114.453, -41.218, -152.325]
  MoveL 8 to (397.22, 170.06, 92.06) mm, rotated rx 122.56 ry -24.48 rz -84.76 deg; joints [67.147, 37.664, -56.735, -114.094, -40.551, -153.434]
  MoveL 9 to (364.46, 170.06, 86.67) mm, rotated rx 122.56 ry -24.48 rz -84.76 deg; joints [68.344, 40.764, -54.654, -113.12, -39.099, -155.989]
  MoveL 10 to (351.69, 170.06, 84.01) mm, rotated rx 122.56 ry -24.48 rz -84.76 deg; joints [68.779, 42.045, -53.848, -112.673, -38.552, -157.016]
  MoveL 11 to (344.57, 170.06, 82.39) mm, rotated rx 122.56 ry -24.48 rz -84.76 deg; joints [69.015, 42.778, -53.398, -112.406, -38.25, -157.599]
  MoveL 12 to (340.58, 170.06, 81.44) mm, rotated rx 122.56 ry -24.48 rz -84.76 deg; joints [69.144, 43.193, -53.146, -112.251, -38.083, -157.928]
  MoveL 13 to (338.06, 170.06, 80.82) mm, rotated rx 122.56 ry -24.48 rz -84.76 deg; joints [69.226, 43.459, -52.986, -112.151, -37.977, -158.138]
  MoveL 14 to (335.56, 170.06, 80.11) mm, rotated rx 122.56 ry -24.48 rz -84.76 deg; joints [69.305, 43.732, -52.837, -112.06, -37.877, -158.333]
  MoveL 15 to (332.95, 170.06, 77.63) mm, rotated rx 122.56 ry -24.48 rz -84.76 deg; joints [69.388, 44.186, -52.849, -112.165, -37.835, -158.284]
  MoveL 16 to (332.4, 170.06, 75.89) mm, rotated rx 122.56 ry -24.48 rz -84.76 deg; joints [69.405, 44.399, -52.97, -112.328, -37.871, -158.096]
  MoveL 17 to (332.35, 170.06, 74.07) mm, rotated rx 122.56 ry -24.48 rz -84.76 deg; joints [69.407, 44.581, -53.142, -112.534, -37.936, -157.836]
  MoveL 18 to (332.35, 170.06, 66.77) mm, rotated rx 122.56 ry -24.48 rz -84.76 deg; joints [69.407, 45.297, -53.846, -113.362, -38.21, -156.784]
  MoveL 19 to (332.35, 170.06, 52.17) mm, rotated rx 122.56 ry -24.48 rz -84.76 deg; joints [69.407, 46.752, -55.228, -114.947, -38.776, -154.759]
  Establecer velocidad (1000.0 mm/s)
  MoveL 20 to (332.35, 170.06, 52.17) mm, rotated rx 122.56 ry -24.48 rz -84.76 deg; joints [69.407, 46.752, -55.228, -114.947, -38.776, -154.759]
  MoveL 21 to (351.96, 170.06, 150.23) mm, rotated rx 122.56 ry -24.48 rz -84.76 deg; joints [68.77, 35.82, -46.815, -103.925, -36.34, -168.011]
  Establecer velocidad (1000.0 mm/s)
  MoveL 22 to (442.77, 170.06, 192.98) mm, rotated rx 122.56 ry -24.48 rz -84.76 deg; joints [65.259, 23.707, -47.429, -101.449, -38.805, -167.89]
  MoveL 23 to (423.16, 170.06, 94.92) mm, rotated rx 122.56 ry -24.48 rz -84.76 deg; joints [66.107, 35.403, -58.417, -114.705, -41.754, -151.456]
  MoveL 24 to (423.16, 170.06, 94.92) mm, rotated rx 122.56 ry -24.48 rz -84.76 deg; joints [66.107, 35.403, -58.417, -114.705, -41.754, -151.456]
  Establecer velocidad (50.0 mm/s)
  MoveL 25 to (441.83, 170.06, 97.34) mm, rotated rx 122.56 ry -24.48 rz -84.76 deg; joints [65.302, 33.756, -59.525, -114.932, -42.596, -150.218]
  MoveL 26 to (460.24, 170.06, 101.28) mm, rotated rx 122.56 ry -24.48 rz -84.76 deg; joints [64.456, 31.96, -60.366, -114.829, -43.334, -149.359]
  MoveL 27 to (478.28, 170.06, 106.75) mm, rotated rx 122.56 ry -24.48 rz -84.76 deg; joints [63.573, 30.004, -60.916, -114.394, -43.957, -148.897]
  MoveL 28 to (495.81, 170.06, 113.69) mm, rotated rx 122.56 ry -24.48 rz -84.76 deg; joints [62.66, 27.886, -61.144, -113.624, -44.454, -148.856]
  MoveL 29 to (517.17, 170.06, 124.58) mm, rotated rx 122.56 ry -24.48 rz -84.76 deg; joints [61.465, 24.951, -60.931, -112.153, -44.904, -149.455]
  MoveL 30 to (537.28, 170.06, 137.67) mm, rotated rx 122.56 ry -24.48 rz -84.76 deg; joints [60.249, 21.758, -60.117, -110.121, -45.169, -150.832]
  MoveL 31 to (555.91, 170.06, 152.79) mm, rotated rx 122.56 ry -24.48 rz -84.76 deg; joints [59.036, 18.335, -58.682, -107.532, -45.29, -153.027]
  MoveL 32 to (572.84, 170.06, 169.77) mm, rotated rx 122.56 ry -24.48 rz -84.76 deg; joints [57.854, 14.737, -56.627, -104.406, -45.333, -156.05]
  Establecer velocidad (1000.0 mm/s)
  MoveL 33 to (572.84, 170.06, 169.77) mm, rotated rx 122.56 ry -24.48 rz -84.76 deg; joints [57.854, 14.737, -56.627, -104.406, -45.333, -156.05]
  MoveL 34 to (592.46, 170.06, 267.83) mm, rotated rx 122.56 ry -24.48 rz -84.76 deg; joints [56.38, 1.916, -40.753, -87.247, -44.682, -178.592]
  Establecer velocidad (1000.0 mm/s)
  MoveL 35 to (713.93, 170.06, 267.83) mm, rotated rx 122.56 ry -24.48 rz -84.76 deg; joints [43.929, -11.111, -39.42, -79.054, -54.29, -178.832]
  MoveL 36 to (694.32, 170.06, 169.77) mm, rotated rx 122.56 ry -24.48 rz -84.76 deg; joints [46.414, 4.341, -59.638, -96.324, -51.808, -153.567]
  MoveL 37 to (694.32, 170.06, 169.77) mm, rotated rx 122.56 ry -24.48 rz -84.76 deg; joints [46.414, 4.341, -59.638, -96.324, -51.808, -153.567]
  Establecer velocidad (50.0 mm/s)
  MoveL 38 to (697.06, 170.06, 153.99) mm, rotated rx 122.56 ry -24.48 rz -84.76 deg; joints [46.081, 6.842, -63.073, -98.666, -52.415, -149.278]
  MoveL 39 to (700.13, 170.06, 138.27) mm, rotated rx 122.56 ry -24.48 rz -84.76 deg; joints [45.701, 9.484, -66.57, -100.919, -53.169, -144.985]
  MoveL 40 to (703.34, 170.06, 122.58) mm, rotated rx 122.56 ry -24.48 rz -84.76 deg; joints [45.299, 12.285, -70.125, -103.086, -54.054, -140.704]
  MoveL 41 to (705.01, 170.06, 107.38) mm, rotated rx 122.56 ry -24.48 rz -84.76 deg; joints [45.088, 15.235, -73.548, -105.241, -54.956, -136.647]
  MoveL 42 to (704.97, 170.06, 92.12) mm, rotated rx 122.56 ry -24.48 rz -84.76 deg; joints [45.094, 18.396, -76.896, -107.462, -55.898, -132.744]
  MoveL 43 to (703.21, 170.06, 77.07) mm, rotated rx 122.56 ry -24.48 rz -84.76 deg; joints [45.316, 21.65, -80.045, -109.675, -56.859, -129.143]
  MoveL 44 to (699.77, 170.06, 62.27) mm, rotated rx 122.56 ry -24.48 rz -84.76 deg; joints [45.747, 24.923, -82.927, -111.844, -57.821, -125.915]
  Establecer velocidad (1000.0 mm/s)
  MoveL 45 to (699.77, 170.06, 62.27) mm, rotated rx 122.56 ry -24.48 rz -84.76 deg; joints [45.747, 24.923, -82.927, -111.844, -57.821, -125.915]
  MoveL 46 to (719.38, 170.06, 160.32) mm, rotated rx 122.56 ry -24.48 rz -84.76 deg; joints [43.201, 3.912, -61.995, -95.184, -53.603, -150.818]

--- program cerlatizqch (robot Fanuc LR Mate 200iD/7L) ---
  Suave(1)
  Establecer velocidad (1000.0 mm/s)
  Est. Ref.: RobotiQ 2F-140 Gripper (Mechanism) Base
  Est. herr: Tool 1
  Mostrar Tool 1
  MoveJ 1 to (226.52, -60.46, 228.77) mm, rotated rx 168.3 ry -14.7 rz -86.98 deg; joints [85.326, 35.729, -18.579, -17.943, -62.565, 103.25]
  MoveL 2 to (226.52, -60.46, 228.77) mm, rotated rx 168.3 ry -14.7 rz -86.98 deg; joints [85.326, 35.729, -18.579, -17.943, -62.565, 103.25]
  MoveL 3 to (206.91, -60.46, 130.71) mm, rotated rx 168.3 ry -14.7 rz -86.98 deg; joints [85.451, 42.635, -27.843, -19.789, -53.759, 106.646]
  MoveL 4 to (206.91, -60.46, 130.71) mm, rotated rx 168.3 ry -14.7 rz -86.98 deg; joints [85.451, 42.635, -27.843, -19.789, -53.759, 106.646]
  Establecer velocidad (50.0 mm/s)
  MoveL 5 to (216.29, -59.67, 130.71) mm, rotated rx 168.3 ry -14.7 rz -86.98 deg; joints [85.33, 41.465, -28.735, -20.032, -52.956, 107.149]
  MoveL 6 to (225.74, -59.68, 130.71) mm, rotated rx 168.3 ry -14.7 rz -86.98 deg; joints [85.27, 40.301, -29.609, -20.271, -52.154, 107.59]
  MoveL 7 to (235.14, -60.49, 130.71) mm, rotated rx 168.3 ry -14.7 rz -86.98 deg; joints [85.273, 39.153, -30.456, -20.503, -51.36, 107.963]
  MoveL 8 to (244.42, -62.09, 130.71) mm, rotated rx 168.3 ry -14.7 rz -86.98 deg; joints [85.341, 38.031, -31.27, -20.726, -50.577, 108.261]
  MoveL 9 to (253.49, -64.46, 131.15) mm, rotated rx 168.3 ry -14.7 rz -86.98 deg; joints [85.476, 36.913, -31.999, -20.923, -49.854, 108.459]
  MoveL 10 to (262.86, -67.6, 132.48) mm, rotated rx 168.3 ry -14.7 rz -86.98 deg; joints [85.678, 35.713, -32.632, -21.089, -49.203, 108.547]
  MoveL 11 to (272.13, -70.38, 134.71) mm, rotated rx 168.3 ry -14.7 rz -86.98 deg; joints [85.855, 34.48, -33.126, -21.219, -48.688, 108.6]
  MoveL 12 to (281.33, -72.64, 137.85) mm, rotated rx 168.3 ry -14.7 rz -86.98 deg; joints [85.993, 33.212, -33.48, -21.314, -48.317, 108.627]
  MoveL 13 to (290.66, -74.45, 140.64) mm, rotated rx 168.3 ry -14.7 rz -86.98 deg; joints [86.095, 31.959, -33.851, -21.421, -47.94, 108.703]
  MoveL 14 to (300.22, -75.82, 142.51) mm, rotated rx 168.3 ry -14.7 rz -86.98 deg; joints [86.16, 30.746, -34.316, -21.567, -47.488, 108.866]
  MoveL 15 to (310.01, -76.73, 143.44) mm, rotated rx 168.3 ry -14.7 rz -86.98 deg; joints [86.182, 29.575, -34.878, -21.756, -46.958, 109.126]
  MoveL 16 to (320.66, -77.15, 143.54) mm, rotated rx 168.3 ry -14.7 rz -86.98 deg; joints [86.155, 28.371, -35.569, -22.002, -46.326, 109.507]
  MoveL 17 to (331.33, -76.98, 143.54) mm, rotated rx 168.3 ry -14.7 rz -86.98 deg; joints [86.073, 27.185, -36.243, -22.259, -45.726, 109.946]
  MoveL 18 to (341.99, -76.98, 143.54) mm, rotated rx 168.3 ry -14.7 rz -86.98 deg; joints [86.003, 26.003, -36.893, -22.512, -45.147, 110.366]
  MoveL 19 to (352.65, -76.98, 143.54) mm, rotated rx 168.3 ry -14.7 rz -86.98 deg; joints [85.931, 24.825, -37.518, -22.763, -44.592, 110.783]
  MoveL 20 to (363.32, -76.98, 143.54) mm, rotated rx 168.3 ry -14.7 rz -86.98 deg; joints [85.856, 23.65, -38.119, -23.012, -44.061, 111.195]
  MoveL 21 to (369.98, -76.98, 143.54) mm, rotated rx 168.3 ry -14.7 rz -86.98 deg; joints [85.808, 22.917, -38.482, -23.166, -43.742, 111.45]
  MoveL 22 to (376.65, -76.98, 143.54) mm, rotated rx 168.3 ry -14.7 rz -86.98 deg; joints [85.759, 22.184, -38.835, -23.319, -43.433, 111.704]
  MoveL 23 to (383.31, -76.98, 143.54) mm, rotated rx 168.3 ry -14.7 rz -86.98 deg; joints [85.709, 21.452, -39.179, -23.471, -43.133, 111.955]
  MoveL 24 to (390.03, -77.17, 143.54) mm, rotated rx 168.3 ry -14.7 rz -86.98 deg; joints [85.677, 20.711, -39.517, -23.62, -42.833, 112.187]
  MoveL 25 to (394.69, -78.33, 143.54) mm, rotated rx 168.3 ry -14.7 rz -86.98 deg; joints [85.76, 20.189, -39.749, -23.71, -42.594, 112.237]
  MoveL 26 to (399.19, -80.59, 143.54) mm, rotated rx 168.3 ry -14.7 rz -86.98 deg; joints [85.964, 19.675, -39.973, -23.782, -42.327, 112.158]
  MoveL 27 to (403.14, -83.9, 143.54) mm, rotated rx 168.3 ry -14.7 rz -86.98 deg; joints [86.286, 19.216, -40.168, -23.828, -42.048, 111.94]
  MoveL 28 to (406.19, -88.02, 143.54) mm, rotated rx 168.3 ry -14.7 rz -86.98 deg; joints [86.705, 18.851, -40.321, -23.841, -41.78, 111.594]
  MoveL 29 to (408.16, -92.59, 143.54) mm, rotated rx 168.3 ry -14.7 rz -86.98 deg; joints [87.183, 18.606, -40.421, -23.823, -41.54, 111.155]
  MoveL 30 to (409.04, -97.21, 143.54) mm, rotated rx 168.3 ry -14.7 rz -86.98 deg; joints [87.675, 18.486, -40.47, -23.776, -41.344, 110.666]
  MoveL 31 to (409.11, -101.66, 143.54) mm, rotated rx 168.3 ry -14.7 rz -86.98 deg; joints [88.155, 18.461, -40.481, -23.711, -41.188, 110.166]
  MoveL 32 to (409.11, -106.11, 143.54) mm, rotated rx 168.3 ry -14.7 rz -86.98 deg; joints [88.634, 18.447, -40.486, -23.643, -41.037, 109.663]
  MoveL 33 to (408.68, -110.65, 143.54) mm, rotated rx 168.3 ry -14.7 rz -86.98 deg; joints [89.124, 18.485, -40.471, -23.56, -40.902, 109.132]
  MoveL 34 to (407.2, -115.28, 143.54) mm, rotated rx 168.3 ry -14.7 rz -86.98 deg; joints [89.624, 18.644, -40.406, -23.451, -40.809, 108.559]
  MoveL 35 to (404.6, -119.64, 143.54) mm, rotated rx 168.3 ry -14.7 rz -86.98 deg; joints [90.093, 18.929, -40.288, -23.32, -40.776, 107.985]
  MoveL 36 to (401.01, -123.35, 143.54) mm, rotated rx 168.3 ry -14.7 rz -86.98 deg; joints [90.486, 19.328, -40.12, -23.178, -40.812, 107.462]
  MoveL 37 to (396.71, -126.09, 143.54) mm, rotated rx 168.3 ry -14.7 rz -86.98 deg; joints [90.771, 19.807, -39.915, -23.036, -40.914, 107.032]
  MoveL 38 to (392.07, -127.73, 143.54) mm, rotated rx 168.3 ry -14.7 rz -86.98 deg; joints [90.935, 20.321, -39.69, -22.906, -41.072, 106.721]
  MoveL 39 to (386, -128.29, 143.54) mm, rotated rx 168.3 ry -14.7 rz -86.98 deg; joints [90.983, 20.992, -39.389, -22.765, -41.335, 106.492]
  MoveL 40 to (380.08, -128.29, 143.54) mm, rotated rx 168.3 ry -14.7 rz -86.98 deg; joints [90.973, 21.645, -39.089, -22.635, -41.616, 106.328]
  MoveL 41 to (374.15, -128.29, 143.54) mm, rotated rx 168.3 ry -14.7 rz -86.98 deg; joints [90.962, 22.298, -38.781, -22.505, -41.903, 106.161]
  MoveL 42 to (368.23, -128.29, 143.54) mm, rotated rx 168.3 ry -14.7 rz -86.98 deg; joints [90.952, 22.951, -38.465, -22.373, -42.198, 105.992]
  MoveL 43 to (362.3, -128.29, 143.54) mm, rotated rx 168.3 ry -14.7 rz -86.98 deg; joints [90.942, 23.604, -38.141, -22.24, -42.5, 105.821]
  MoveL 44 to (356.38, -128.29, 143.54) mm, rotated rx 168.3 ry -14.7 rz -86.98 deg; joints [90.933, 24.258, -37.81, -22.106, -42.81, 105.647]
  MoveL 45 to (344.65, -128.29, 143.54) mm, rotated rx 168.3 ry -14.7 rz -86.98 deg; joints [90.914, 25.555, -37.133, -21.839, -43.444, 105.296]
  MoveL 46 to (332.92, -128.29, 143.54) mm, rotated rx 168.3 ry -14.7 rz -86.98 deg; joints [90.896, 26.857, -36.425, -21.569, -44.106, 104.937]
  MoveL 47 to (321.2, -128.68, 143.54) mm, rotated rx 168.3 ry -14.7 rz -86.98 deg; joints [90.916, 28.165, -35.687, -21.29, -44.788, 104.531]
  MoveL 48 to (309.53, -129.88, 143.41) mm, rotated rx 168.3 ry -14.7 rz -86.98 deg; joints [91.006, 29.484, -34.935, -21.004, -45.462, 104.051]
  MoveL 49 to (299.82, -131.49, 142.45) mm, rotated rx 168.3 ry -14.7 rz -86.98 deg; joints [91.135, 30.646, -34.385, -20.789, -45.938, 103.639]
  MoveL 50 to (290.35, -133.62, 140.57) mm, rotated rx 168.3 ry -14.7 rz -86.98 deg; joints [91.306, 31.847, -33.933, -20.604, -46.311, 103.233]
  MoveL 51 to (281.11, -136.13, 137.77) mm, rotated rx 168.3 ry -14.7 rz -86.98 deg; joints [91.506, 33.084, -33.574, -20.448, -46.589, 102.845]
  MoveL 52 to (271.92, -138.27, 134.65) mm, rotated rx 168.3 ry -14.7 rz -86.98 deg; joints [91.669, 34.341, -33.228, -20.304, -46.866, 102.504]
  MoveL 53 to (262.48, -139.96, 132.41) mm, rotated rx 168.3 ry -14.7 rz -86.98 deg; joints [91.788, 35.576, -32.736, -20.124, -47.293, 102.144]
  MoveL 54 to (252.81, -141.17, 131.08) mm, rotated rx 168.3 ry -14.7 rz -86.98 deg; joints [91.863, 36.788, -32.096, -19.909, -47.873, 101.766]
  MoveL 55 to (243.98, -141.82, 130.71) mm, rotated rx 168.3 ry -14.7 rz -86.98 deg; joints [91.893, 37.855, -31.395, -19.691, -48.524, 101.416]
  MoveL 56 to (235.07, -142.04, 130.71) mm, rotated rx 168.3 ry -14.7 rz -86.98 deg; joints [91.887, 38.92, -30.626, -19.467, -49.251, 101.081]
  MoveL 57 to (226.16, -142.04, 130.71) mm, rotated rx 168.3 ry -14.7 rz -86.98 deg; joints [91.863, 39.999, -29.833, -19.248, -50.006, 100.761]
  MoveL 58 to (217.26, -141.56, 130.71) mm, rotated rx 168.3 ry -14.7 rz -86.98 deg; joints [91.802, 41.091, -29.017, -19.039, -50.794, 100.479]
  MoveL 59 to (208.48, -140.06, 130.71) mm, rotated rx 168.3 ry -14.7 rz -86.98 deg; joints [91.663, 42.184, -28.188, -18.849, -51.617, 100.282]
  MoveL 60 to (199.93, -137.56, 130.87) mm, rotated rx 168.3 ry -14.7 rz -86.98 deg; joints [91.45, 43.254, -27.341, -18.676, -52.48, 100.162]
  MoveL 61 to (191.78, -134.11, 131.41) mm, rotated rx 168.3 ry -14.7 rz -86.98 deg; joints [91.171, 44.273, -26.468, -18.517, -53.387, 100.109]
  MoveL 62 to (184.04, -129.74, 132.28) mm, rotated rx 168.3 ry -14.7 rz -86.98 deg; joints [90.828, 45.242, -25.577, -18.375, -54.329, 100.123]
  MoveL 63 to (176.91, -124.55, 133.38) mm, rotated rx 168.3 ry -14.7 rz -86.98 deg; joints [90.431, 46.141, -24.701, -18.253, -55.274, 100.203]
  MoveL 64 to (172.96, -121.08, 134.12) mm, rotated rx 168.3 ry -14.7 rz -86.98 deg; joints [90.169, 46.645, -24.189, -18.19, -55.835, 100.283]
  MoveL 65 to (169.24, -117.34, 134.9) mm, rotated rx 168.3 ry -14.7 rz -86.98 deg; joints [89.89, 47.123, -23.691, -18.135, -56.388, 100.388]
  MoveL 66 to (165.8, -113.31, 135.7) mm, rotated rx 168.3 ry -14.7 rz -86.98 deg; joints [89.593, 47.572, -23.212, -18.089, -56.927, 100.521]
  MoveL 67 to (163.23, -108.67, 136.34) mm, rotated rx 168.3 ry -14.7 rz -86.98 deg; joints [89.252, 47.913, -22.843, -18.074, -57.376, 100.739]
  MoveL 68 to (161.89, -103.51, 136.69) mm, rotated rx 168.3 ry -14.7 rz -86.98 deg; joints [88.874, 48.1, -22.64, -18.099, -57.677, 101.057]
  MoveL 69 to (161.72, -97.55, 136.74) mm, rotated rx 168.3 ry -14.7 rz -86.98 deg; joints [88.436, 48.143, -22.599, -18.165, -57.842, 101.496]
  MoveL 70 to (162.18, -91.62, 136.62) mm, rotated rx 168.3 ry -14.7 rz -86.98 deg; joints [87.998, 48.108, -22.645, -18.247, -57.925, 101.967]
  MoveL 71 to (163.69, -85.89, 136.22) mm, rotated rx 168.3 ry -14.7 rz -86.98 deg; joints [87.572, 47.942, -22.836, -18.354, -57.866, 102.478]
  MoveL 72 to (166.18, -80.56, 135.61) mm, rotated rx 168.3 ry -14.7 rz -86.98 deg; joints [87.171, 47.653, -23.16, -18.482, -57.675, 103.013]
  MoveL 73 to (169.57, -75.75, 134.83) mm, rotated rx 168.3 ry -14.7 rz -86.98 deg; joints [86.802, 47.248, -23.6, -18.629, -57.366, 103.56]
  MoveL 74 to (173.74, -71.64, 133.97) mm, rotated rx 168.3 ry -14.7 rz -86.98 deg; joints [86.478, 46.744, -24.132, -18.79, -56.957, 104.096]
  MoveL 75 to (178.57, -68.32, 133.09) mm, rotated rx 168.3 ry -14.7 rz -86.98 deg; joints [86.208, 46.153, -24.733, -18.958, -56.468, 104.608]
  MoveL 76 to (183.92, -65.91, 132.29) mm, rotated rx 168.3 ry -14.7 rz -86.98 deg; joints [85.999, 45.493, -25.376, -19.13, -55.922, 105.075]
  MoveL 77 to (189.54, -64.09, 131.63) mm, rotated rx 168.3 ry -14.7 rz -86.98 deg; joints [85.831, 44.796, -26.025, -19.301, -55.359, 105.507]
  MoveL 78 to (195.25, -62.58, 131.14) mm, rotated rx 168.3 ry -14.7 rz -86.98 deg; joints [85.684, 44.089, -26.653, -19.468, -54.811, 105.913]
  MoveL 79 to (201.04, -61.36, 130.83) mm, rotated rx 168.3 ry -14.7 rz -86.98 deg; joints [85.557, 43.369, -27.259, -19.631, -54.277, 106.293]
  MoveL 80 to (206.91, -60.46, 130.71) mm, rotated rx 168.3 ry -14.7 rz -86.98 deg; joints [85.451, 42.635, -27.843, -19.789, -53.759, 106.646]
  Establecer velocidad (1000.0 mm/s)
  MoveL 81 to (206.91, -60.46, 130.71) mm, rotated rx 168.3 ry -14.7 rz -86.98 deg; joints [85.451, 42.635, -27.843, -19.789, -53.759, 106.646]
  MoveL 82 to (226.52, -60.46, 228.77) mm, rotated rx 168.3 ry -14.7 rz -86.98 deg; joints [85.326, 35.729, -18.579, -17.943, -62.565, 103.25]
  Establecer velocidad (1000.0 mm/s)
  MoveL 83 to (379.58, -128.44, 281) mm, rotated rx 168.3 ry -14.7 rz -86.98 deg; joints [90.986, 13.982, -21.049, -17.423, -58.594, 98.287]
  MoveL 84 to (359.97, -128.44, 182.94) mm, rotated rx 168.3 ry -14.7 rz -86.98 deg; joints [90.953, 21.212, -33.011, -20.366, -47.278, 103.169]
  MoveL 85 to (359.97, -128.44, 182.94) mm, rotated rx 168.3 ry -14.7 rz -86.98 deg; joints [90.953, 21.212, -33.011, -20.366, -47.278, 103.169]
  Establecer velocidad (50.0 mm/s)
  MoveL 86 to (376.1, -127.67, 182.94) mm, rotated rx 168.3 ry -14.7 rz -86.98 deg; joints [90.902, 19.348, -33.78, -20.626, -46.572, 103.592]
  MoveL 87 to (392.1, -125.43, 182.94) mm, rotated rx 168.3 ry -14.7 rz -86.98 deg; joints [90.695, 17.494, -34.482, -20.902, -45.977, 104.159]
  MoveL 88 to (397.3, -123.99, 182.94) mm, rotated rx 168.3 ry -14.7 rz -86.98 deg; joints [90.549, 16.891, -34.696, -21.002, -45.82, 104.421]
  MoveL 89 to (402.02, -121.44, 182.94) mm, rotated rx 168.3 ry -14.7 rz -86.98 deg; joints [90.283, 16.341, -34.886, -21.115, -45.722, 104.801]
  MoveL 90 to (406.11, -117.92, 182.94) mm, rotated rx 168.3 ry -14.7 rz -86.98 deg; joints [89.908, 15.866, -35.045, -21.236, -45.684, 105.282]
  MoveL 91 to (409.3, -113.58, 182.94) mm, rotated rx 168.3 ry -14.7 rz -86.98 deg; joints [89.439, 15.498, -35.166, -21.358, -45.711, 105.843]
  MoveL 92 to (411.27, -108.57, 182.94) mm, rotated rx 168.3 ry -14.7 rz -86.98 deg; joints [88.895, 15.278, -35.236, -21.472, -45.807, 106.456]
  MoveL 93 to (411.78, -103.25, 182.94) mm, rotated rx 168.3 ry -14.7 rz -86.98 deg; joints [88.317, 15.233, -35.25, -21.569, -45.967, 107.075]
  MoveL 94 to (411.63, -98.97, 182.94) mm, rotated rx 168.3 ry -14.7 rz -86.98 deg; joints [87.855, 15.267, -35.24, -21.637, -46.117, 107.557]
  MoveL 95 to (410.65, -94.86, 182.94) mm, rotated rx 168.3 ry -14.7 rz -86.98 deg; joints [87.415, 15.4, -35.197, -21.689, -46.289, 107.998]
  MoveL 96 to (408.85, -91.01, 182.94) mm, rotated rx 168.3 ry -14.7 rz -86.98 deg; joints [87.009, 15.632, -35.122, -21.722, -46.481, 108.386]
  MoveL 97 to (406.34, -87.61, 182.94) mm, rotated rx 168.3 ry -14.7 rz -86.98 deg; joints [86.66, 15.945, -35.019, -21.737, -46.682, 108.698]
  MoveL 98 to (403.26, -84.69, 182.94) mm, rotated rx 168.3 ry -14.7 rz -86.98 deg; joints [86.368, 16.321, -34.893, -21.734, -46.888, 108.939]
  MoveL 99 to (398.55, -81.71, 182.94) mm, rotated rx 168.3 ry -14.7 rz -86.98 deg; joints [86.086, 16.889, -34.697, -21.707, -47.156, 109.135]
  MoveL 100 to (393.23, -79.95, 182.94) mm, rotated rx 168.3 ry -14.7 rz -86.98 deg; joints [85.94, 17.517, -34.474, -21.651, -47.408, 109.174]
  MoveL 101 to (387.71, -79.03, 182.94) mm, rotated rx 168.3 ry -14.7 rz -86.98 deg; joints [85.886, 18.161, -34.237, -21.578, -47.645, 109.112]
  MoveL 102 to (382.16, -78.28, 182.94) mm, rotated rx 168.3 ry -14.7 rz -86.98 deg; joints [85.85, 18.807, -33.992, -21.501, -47.884, 109.028]
  MoveL 103 to (376.6, -77.7, 182.94) mm, rotated rx 168.3 ry -14.7 rz -86.98 deg; joints [85.832, 19.453, -33.739, -21.42, -48.124, 108.922]
  MoveL 104 to (371.01, -77.29, 182.94) mm, rotated rx 168.3 ry -14.7 rz -86.98 deg; joints [85.831, 20.1, -33.478, -21.336, -48.368, 108.795]
  MoveL 105 to (357.83, -76.95, 182.94) mm, rotated rx 168.3 ry -14.7 rz -86.98 deg; joints [85.892, 21.623, -32.834, -21.122, -48.949, 108.422]
  MoveL 106 to (344.64, -77.42, 182.94) mm, rotated rx 168.3 ry -14.7 rz -86.98 deg; joints [86.027, 23.142, -32.152, -20.892, -49.545, 107.958]
  MoveL 107 to (336.87, -78.26, 182.94) mm, rotated rx 168.3 ry -14.7 rz -86.98 deg; joints [86.158, 24.035, -31.733, -20.747, -49.898, 107.627]
  MoveL 108 to (329.21, -79.58, 182.94) mm, rotated rx 168.3 ry -14.7 rz -86.98 deg; joints [86.328, 24.915, -31.307, -20.597, -50.245, 107.253]
  MoveL 109 to (321.57, -80.78, 182.94) mm, rotated rx 168.3 ry -14.7 rz -86.98 deg; joints [86.485, 25.796, -30.867, -20.447, -50.61, 106.891]
  MoveL 110 to (313.81, -80.7, 182.94) mm, rotated rx 168.3 ry -14.7 rz -86.98 deg; joints [86.52, 26.704, -30.401, -20.309, -51.036, 106.645]
  MoveL 111 to (306.05, -80.58, 182.94) mm, rotated rx 168.3 ry -14.7 rz -86.98 deg; joints [86.552, 27.616, -29.92, -20.171, -51.478, 106.399]
  MoveL 112 to (298.3, -80.59, 182.94) mm, rotated rx 168.3 ry -14.7 rz -86.98 deg; joints [86.595, 28.532, -29.424, -20.03, -51.931, 106.137]
  MoveL 113 to (294.77, -80.7, 182.94) mm, rotated rx 168.3 ry -14.7 rz -86.98 deg; joints [86.623, 28.949, -29.194, -19.964, -52.139, 106.008]
  MoveL 114 to (291.25, -80.91, 182.94) mm, rotated rx 168.3 ry -14.7 rz -86.98 deg; joints [86.659, 29.366, -28.961, -19.897, -52.347, 105.87]
  MoveL 115 to (287.74, -81.26, 182.94) mm, rotated rx 168.3 ry -14.7 rz -86.98 deg; joints [86.707, 29.782, -28.726, -19.829, -52.553, 105.719]
  MoveL 116 to (284.32, -82.1, 182.94) mm, rotated rx 168.3 ry -14.7 rz -86.98 deg; joints [86.798, 30.186, -28.496, -19.755, -52.743, 105.527]
  MoveL 117 to (281.45, -84.14, 182.94) mm, rotated rx 168.3 ry -14.7 rz -86.98 deg; joints [86.989, 30.517, -28.305, -19.677, -52.866, 105.248]
  MoveL 118 to (279.68, -86.5, 182.94) mm, rotated rx 168.3 ry -14.7 rz -86.98 deg; joints [87.201, 30.715, -28.19, -19.615, -52.911, 104.978]
  MoveL 119 to (278.72, -89.28, 182.94) mm, rotated rx 168.3 ry -14.7 rz -86.98 deg; joints [87.445, 30.816, -28.132, -19.562, -52.894, 104.699]
  MoveL 120 to (278.78, -92.22, 182.94) mm, rotated rx 168.3 ry -14.7 rz -86.98 deg; joints [87.699, 30.793, -28.145, -19.526, -52.807, 104.44]
  MoveL 121 to (280.1, -96.44, 182.94) mm, rotated rx 168.3 ry -14.7 rz -86.98 deg; joints [88.06, 30.615, -28.248, -19.494, -52.603, 104.107]
  MoveL 122 to (281.55, -100.62, 182.94) mm, rotated rx 168.3 ry -14.7 rz -86.98 deg; joints [88.419, 30.426, -28.358, -19.464, -52.395, 103.777]
  MoveL 123 to (281.1, -102.5, 182.94) mm, rotated rx 168.3 ry -14.7 rz -86.98 deg; joints [88.583, 30.473, -28.33, -19.43, -52.373, 103.593]
  MoveL 124 to (280.55, -104.38, 182.94) mm, rotated rx 168.3 ry -14.7 rz -86.98 deg; joints [88.748, 30.535, -28.295, -19.393, -52.358, 103.406]
  MoveL 125 to (280.01, -106.27, 182.94) mm, rotated rx 168.3 ry -14.7 rz -86.98 deg; joints [88.913, 30.595, -28.26, -19.356, -52.343, 103.218]
  MoveL 126 to (279.47, -108.16, 182.94) mm, rotated rx 168.3 ry -14.7 rz -86.98 deg; joints [89.078, 30.656, -28.225, -19.32, -52.328, 103.03]
  MoveL 127 to (278.95, -110.06, 182.94) mm, rotated rx 168.3 ry -14.7 rz -86.98 deg; joints [89.243, 30.715, -28.19, -19.283, -52.312, 102.842]
  MoveL 128 to (278.65, -111.99, 182.94) mm, rotated rx 168.3 ry -14.7 rz -86.98 deg; joints [89.41, 30.749, -28.171, -19.249, -52.282, 102.658]
  MoveL 129 to (279.11, -115.84, 182.94) mm, rotated rx 168.3 ry -14.7 rz -86.98 deg; joints [89.743, 30.69, -28.204, -19.2, -52.153, 102.322]
  MoveL 130 to (280.8, -119.34, 182.94) mm, rotated rx 168.3 ry -14.7 rz -86.98 deg; joints [90.047, 30.486, -28.323, -19.178, -51.954, 102.051]
  MoveL 131 to (283.36, -122.25, 182.94) mm, rotated rx 168.3 ry -14.7 rz -86.98 deg; joints [90.301, 30.18, -28.499, -19.178, -51.714, 101.856]
  MoveL 132 to (286.74, -124.16, 182.94) mm, rotated rx 168.3 ry -14.7 rz -86.98 deg; joints [90.47, 29.777, -28.729, -19.208, -51.448, 101.774]
  MoveL 133 to (290.57, -124.79, 182.94) mm, rotated rx 168.3 ry -14.7 rz -86.98 deg; joints [90.529, 29.319, -28.987, -19.265, -51.188, 101.82]
  MoveL 134 to (294.45, -125.15, 182.94) mm, rotated rx 168.3 ry -14.7 rz -86.98 deg; joints [90.563, 28.858, -29.244, -19.328, -50.935, 101.892]
  MoveL 135 to (298.34, -125.32, 182.94) mm, rotated rx 168.3 ry -14.7 rz -86.98 deg; joints [90.582, 28.397, -29.498, -19.393, -50.69, 101.981]
  MoveL 136 to (302.23, -125.36, 182.94) mm, rotated rx 168.3 ry -14.7 rz -86.98 deg; joints [90.59, 27.936, -29.748, -19.46, -50.452, 102.081]
  MoveL 137 to (306.13, -125.32, 182.94) mm, rotated rx 168.3 ry -14.7 rz -86.98 deg; joints [90.589, 27.476, -29.994, -19.528, -50.22, 102.188]
  MoveL 138 to (310.49, -125.2, 182.94) mm, rotated rx 168.3 ry -14.7 rz -86.98 deg; joints [90.583, 26.963, -30.266, -19.605, -49.966, 102.313]
  MoveL 139 to (314.85, -125.06, 182.94) mm, rotated rx 168.3 ry -14.7 rz -86.98 deg; joints [90.574, 26.451, -30.532, -19.683, -49.718, 102.44]
  MoveL 140 to (319.21, -124.92, 182.94) mm, rotated rx 168.3 ry -14.7 rz -86.98 deg; joints [90.565, 25.94, -30.794, -19.759, -49.474, 102.566]
  MoveL 141 to (323.57, -124.82, 182.94) mm, rotated rx 168.3 ry -14.7 rz -86.98 deg; joints [90.56, 25.43, -31.051, -19.835, -49.233, 102.685]
  MoveL 142 to (327.85, -125.65, 182.94) mm, rotated rx 168.3 ry -14.7 rz -86.98 deg; joints [90.641, 24.931, -31.298, -19.893, -48.977, 102.71]
  MoveL 143 to (332.17, -126.69, 182.94) mm, rotated rx 168.3 ry -14.7 rz -86.98 deg; joints [90.744, 24.43, -31.543, -19.948, -48.717, 102.711]
  MoveL 144 to (336.92, -127.76, 182.94) mm, rotated rx 168.3 ry -14.7 rz -86.98 deg; joints [90.852, 23.88, -31.806, -20.008, -48.438, 102.717]
  MoveL 145 to (340.7, -128.25, 182.94) mm, rotated rx 168.3 ry -14.7 rz -86.98 deg; joints [90.904, 23.443, -32.012, -20.061, -48.23, 102.755]
  MoveL 146 to (343.65, -128.42, 182.94) mm, rotated rx 168.3 ry -14.7 rz -86.98 deg; joints [90.924, 23.1, -32.171, -20.106, -48.075, 102.807]
  MoveL 147 to (346.41, -128.44, 182.94) mm, rotated rx 168.3 ry -14.7 rz -86.98 deg; joints [90.931, 22.781, -32.317, -20.15, -47.935, 102.867]
  MoveL 148 to (348.8, -128.44, 182.94) mm, rotated rx 168.3 ry -14.7 rz -86.98 deg; joints [90.935, 22.503, -32.443, -20.189, -47.816, 102.922]
  MoveL 149 to (351.88, -128.44, 182.94) mm, rotated rx 168.3 ry -14.7 rz -86.98 deg; joints [90.94, 22.147, -32.603, -20.238, -47.665, 102.991]
  MoveL 150 to (355.74, -128.44, 182.94) mm, rotated rx 168.3 ry -14.7 rz -86.98 deg; joints [90.946, 21.701, -32.8, -20.299, -47.478, 103.077]
  MoveL 151 to (359.97, -128.44, 182.94) mm, rotated rx 168.3 ry -14.7 rz -86.98 deg; joints [90.953, 21.212, -33.011, -20.366, -47.278, 103.169]
  Establecer velocidad (1000.0 mm/s)
  MoveL 152 to (359.97, -128.44, 182.94) mm, rotated rx 168.3 ry -14.7 rz -86.98 deg; joints [90.953, 21.212, -33.011, -20.366, -47.278, 103.169]
  MoveL 153 to (379.58, -128.44, 281) mm, rotated rx 168.3 ry -14.7 rz -86.98 deg; joints [90.986, 13.982, -21.049, -17.423, -58.594, 98.287]

